screen "P_GraphicView_1" 1280x800
   GraphicView "Default" at 10,10 size 100x60
   TextField "Label_Default" at 10,72 size 108x16; Text 'Default'
   GraphicView "BackColor" at 120,10 size 100x60
   TextField "Label_BackColor" at 120,72 size 108x16; Text 'BackColor'
   GraphicView "BackFillStyle" at 230,10 size 100x60
   TextField "Label_BackFillStyle" at 230,72 size 108x16; Text 'BackFillStyle'
   GraphicView "BorderColor" at 340,10 size 100x60
   TextField "Label_BorderColor" at 340,72 size 108x16; Text 'BorderColor'
   GraphicView "BorderWidth" at 450,10 size 100x60
   TextField "Label_BorderWidth" at 450,72 size 108x16; Text 'BorderWidth'
   GraphicView "EdgeStyle" at 560,10 size 100x60
   TextField "Label_EdgeStyle" at 560,72 size 108x16; Text 'EdgeStyle'
   GraphicView "EdgeStyle_2" at 670,10 size 100x60
   TextField "Label_EdgeStyle_2" at 670,72 size 108x16; Text 'EdgeStyle_2'
   GraphicView "EdgeStyle_3" at 780,10 size 100x60
   TextField "Label_EdgeStyle_3" at 780,72 size 108x16; Text 'EdgeStyle_3'
   GraphicView "EdgeStyle_4" at 890,10 size 100x60
   TextField "Label_EdgeStyle_4" at 890,72 size 108x16; Text 'EdgeStyle_4'
   GraphicView "FitToLargest" at 1000,10 size 100x60
   TextField "Label_FitToLargest" at 1000,72 size 108x16; Text 'FitToLargest'
   GraphicView "Flashing" at 1110,10 size 100x60
   TextField "Label_Flashing" at 1110,72 size 108x16; Text 'Flashing'
   GraphicView "TransparentColor" at 10,96 size 100x60
   TextField "Label_TransparentColor" at 10,158 size 108x16; Text 'TransparentColor'
   GraphicView "UseTransparentColor" at 120,96 size 100x60
   TextField "Label_UseTransparentColor" at 120,158 size 108x16; Text 'UseTransparentColor'
   Button "Next" at 1238,776 size 40x22; TextOff 'Text'
      on Click: ActivateScreen("P_IOField_1", 0)

screen "P_IOField_1" 1280x800
   IOField "Default" at 10,10 size 100x30
   TextField "Label_Default" at 10,42 size 108x16; Text 'Default'
   IOField "AboveUpperLimitColor" at 120,10 size 100x30
   TextField "Label_AboveUpperLimitColor" at 120,42 size 108x16; Text 'AboveUpperLimitColor'
   IOField "BackColor" at 230,10 size 100x30
   TextField "Label_BackColor" at 230,42 size 108x16; Text 'BackColor'
   IOField "BackFillStyle" at 340,10 size 100x30
   TextField "Label_BackFillStyle" at 340,42 size 108x16; Text 'BackFillStyle'
   IOField "BelowLowerLimitColor" at 450,10 size 100x30
   TextField "Label_BelowLowerLimitColor" at 450,42 size 108x16; Text 'BelowLowerLimitColor'
   IOField "BorderBackColor" at 560,10 size 100x30
   TextField "Label_BorderBackColor" at 560,42 size 108x16; Text 'BorderBackColor'
   IOField "BorderColor" at 670,10 size 100x30
   TextField "Label_BorderColor" at 670,42 size 108x16; Text 'BorderColor'
   IOField "BorderWidth" at 780,10 size 100x30
   TextField "Label_BorderWidth" at 780,42 size 108x16; Text 'BorderWidth'
   IOField "BottomMargin" at 890,10 size 100x30
   TextField "Label_BottomMargin" at 890,42 size 108x16; Text 'BottomMargin'
   IOField "CornerRadius" at 1000,10 size 100x30
   TextField "Label_CornerRadius" at 1000,42 size 108x16; Text 'CornerRadius'
   IOField "DataFormat_3" at 1110,10 size 100x30
   TextField "Label_DataFormat_3" at 1110,42 size 108x16; Text 'DataFormat_3'
   IOField "EdgeStyle" at 10,66 size 100x30
   TextField "Label_EdgeStyle" at 10,98 size 108x16; Text 'EdgeStyle'
   IOField "EdgeStyle_2" at 120,66 size 100x30
   TextField "Label_EdgeStyle_2" at 120,98 size 108x16; Text 'EdgeStyle_2'
   IOField "EdgeStyle_3" at 230,66 size 100x30
   TextField "Label_EdgeStyle_3" at 230,98 size 108x16; Text 'EdgeStyle_3'
   IOField "EdgeStyle_4" at 340,66 size 100x30
   TextField "Label_EdgeStyle_4" at 340,98 size 108x16; Text 'EdgeStyle_4'
   IOField "FieldLength" at 450,66 size 100x30
   TextField "Label_FieldLength" at 450,98 size 108x16; Text 'FieldLength'
   IOField "FitToLargest" at 560,66 size 100x30
   TextField "Label_FitToLargest" at 560,98 size 108x16; Text 'FitToLargest'
   IOField "Flashing" at 670,66 size 100x30
   TextField "Label_Flashing" at 670,98 size 108x16; Text 'Flashing'
   IOField "ForeColor" at 780,66 size 100x30
   TextField "Label_ForeColor" at 780,98 size 108x16; Text 'ForeColor'
   IOField "FormatPattern" at 890,66 size 100x30; FormatPattern 99.9
   TextField "Label_FormatPattern" at 890,98 size 108x16; Text 'FormatPattern'
   IOField "HorizontalAlignment" at 1000,66 size 100x30
   TextField "Label_HorizontalAlignment" at 1000,98 size 108x16; Text 'HorizontalAlignment'
   IOField "HorizontalAlignment_2" at 1110,66 size 100x30
   TextField "Label_HorizontalAlignment_2" at 1110,98 size 108x16; Text 'HorizontalAlignment_2'
   IOField "LeftMargin" at 10,122 size 100x30
   TextField "Label_LeftMargin" at 10,154 size 108x16; Text 'LeftMargin'
   IOField "Mode" at 120,122 size 100x30
   TextField "Label_Mode" at 120,154 size 108x16; Text 'Mode'
   IOField "Mode_2" at 230,122 size 100x30
   TextField "Label_Mode_2" at 230,154 size 108x16; Text 'Mode_2'
   IOField "RightMargin" at 340,122 size 100x30
   TextField "Label_RightMargin" at 340,154 size 108x16; Text 'RightMargin'
   IOField "ShiftDecimalPoint" at 450,122 size 100x30
   TextField "Label_ShiftDecimalPoint" at 450,154 size 108x16; Text 'ShiftDecimalPoint'
   IOField "ShowLeadingZeros" at 560,122 size 100x30
   TextField "Label_ShowLeadingZeros" at 560,154 size 108x16; Text 'ShowLeadingZeros'
   IOField "TopMargin" at 670,122 size 100x30
   TextField "Label_TopMargin" at 670,154 size 108x16; Text 'TopMargin'
   IOField "Unit" at 780,122 size 100x30; Unit mm
   TextField "Label_Unit" at 780,154 size 108x16; Text 'Unit'
   IOField "UseDesignColorSchema" at 890,122 size 100x30
   TextField "Label_UseDesignColorSchema" at 890,154 size 108x16; Text 'UseDesignColorSchema'
   IOField "VerticalAlignment" at 1000,122 size 100x30
   TextField "Label_VerticalAlignment" at 1000,154 size 108x16; Text 'VerticalAlignment'
   IOField "VerticalAlignment_2" at 1110,122 size 100x30
   TextField "Label_VerticalAlignment_2" at 1110,154 size 108x16; Text 'VerticalAlignment_2'
   Button "Next" at 1238,776 size 40x22; TextOff 'Text'
      on Click: ActivateScreen("P_Button_1", 0)

screen "P_Button_1" 1280x800
   Button "Default" at 10,10 size 100x40; TextOff 'Text'
   TextField "Label_Default" at 10,52 size 108x16; Text 'Default'
   Button "BackColor" at 120,10 size 100x40; TextOff 'Text'
   TextField "Label_BackColor" at 120,52 size 108x16; Text 'BackColor'
   Button "BackFillStyle" at 230,10 size 100x40; TextOff 'Text'
   TextField "Label_BackFillStyle" at 230,52 size 108x16; Text 'BackFillStyle'
   Button "BorderBackColor" at 340,10 size 100x40; TextOff 'Text'
   TextField "Label_BorderBackColor" at 340,52 size 108x16; Text 'BorderBackColor'
   Button "BorderColor" at 450,10 size 100x40; TextOff 'Text'
   TextField "Label_BorderColor" at 450,52 size 108x16; Text 'BorderColor'
   Button "BorderWidth" at 560,10 size 100x40; TextOff 'Text'
   TextField "Label_BorderWidth" at 560,52 size 108x16; Text 'BorderWidth'
   Button "CornerRadius" at 670,10 size 100x40; TextOff 'Text'
   TextField "Label_CornerRadius" at 670,52 size 108x16; Text 'CornerRadius'
   Button "EdgeStyle" at 780,10 size 100x40; TextOff 'Text'
   TextField "Label_EdgeStyle" at 780,52 size 108x16; Text 'EdgeStyle'
   Button "EdgeStyle_2" at 890,10 size 100x40; TextOff 'Text'
   TextField "Label_EdgeStyle_2" at 890,52 size 108x16; Text 'EdgeStyle_2'
   Button "EdgeStyle_3" at 1000,10 size 100x40; TextOff 'Text'
   TextField "Label_EdgeStyle_3" at 1000,52 size 108x16; Text 'EdgeStyle_3'
   Button "EdgeStyle_4" at 1110,10 size 100x40; TextOff 'Text'
   TextField "Label_EdgeStyle_4" at 1110,52 size 108x16; Text 'EdgeStyle_4'
   Button "FirstGradientColor" at 10,76 size 100x40; TextOff 'Text'
   TextField "Label_FirstGradientColor" at 10,118 size 108x16; Text 'FirstGradientColor'
   Button "FirstGradientOffset" at 120,76 size 100x40; TextOff 'Text'
   TextField "Label_FirstGradientOffset" at 120,118 size 108x16; Text 'FirstGradientOffset'
   Button "FitToLargest" at 230,76 size 100x40; TextOff 'Text'
   TextField "Label_FitToLargest" at 230,118 size 108x16; Text 'FitToLargest'
   Button "Flashing" at 340,76 size 100x40; TextOff 'Text'
   TextField "Label_Flashing" at 340,118 size 108x16; Text 'Flashing'
   Button "FocusColor" at 450,76 size 100x40; TextOff 'Text'
   TextField "Label_FocusColor" at 450,118 size 108x16; Text 'FocusColor'
   Button "FocusWidth" at 560,76 size 100x40; TextOff 'Text'
   TextField "Label_FocusWidth" at 560,118 size 108x16; Text 'FocusWidth'
   Button "ForeColor" at 670,76 size 100x40; TextOff 'Text'
   TextField "Label_ForeColor" at 670,118 size 108x16; Text 'ForeColor'
   Button "HorizontalAlignment" at 780,76 size 100x40; TextOff 'Text'
   TextField "Label_HorizontalAlignment" at 780,118 size 108x16; Text 'HorizontalAlignment'
   Button "HorizontalAlignment_2" at 890,76 size 100x40; TextOff 'Text'
   TextField "Label_HorizontalAlignment_2" at 890,118 size 108x16; Text 'HorizontalAlignment_2'
   Button "HorizontalPictureAlignment" at 1000,76 size 100x40; TextOff 'Text'
   TextField "Label_HorizontalPictureAlignment" at 1000,118 size 108x16; Text 'HorizontalPictureAlignment'
   Button "HorizontalPictureAlignment_2" at 1110,76 size 100x40; TextOff 'Text'
   TextField "Label_HorizontalPictureAlignment_2" at 1110,118 size 108x16; Text 'HorizontalPictureAlignment_2'
   Button "MiddleGradientColor" at 10,142 size 100x40; TextOff 'Text'
   TextField "Label_MiddleGradientColor" at 10,184 size 108x16; Text 'MiddleGradientColor'
   Button "Mode_5" at 120,142 size 100x40; TextOff 'Text'
   TextField "Label_Mode_5" at 120,184 size 108x16; Text 'Mode_5'
   Button "Mode_7" at 230,142 size 100x40; TextOff 'Text'
   TextField "Label_Mode_7" at 230,184 size 108x16; Text 'Mode_7'
   Button "PictureAreaBottomMargin" at 340,142 size 100x40; TextOff 'Text'
   TextField "Label_PictureAreaBottomMargin" at 340,184 size 108x16; Text 'PictureAreaBottomMargin'
   Button "PictureAreaLeftMargin" at 450,142 size 100x40; TextOff 'Text'
   TextField "Label_PictureAreaLeftMargin" at 450,184 size 108x16; Text 'PictureAreaLeftMargin'
   Button "PictureAreaRightMargin" at 560,142 size 100x40; TextOff 'Text'
   TextField "Label_PictureAreaRightMargin" at 560,184 size 108x16; Text 'PictureAreaRightMargin'
   Button "PictureAreaTopMargin" at 670,142 size 100x40; TextOff 'Text'
   TextField "Label_PictureAreaTopMargin" at 670,184 size 108x16; Text 'PictureAreaTopMargin'
   Button "SecondGradientColor" at 780,142 size 100x40; TextOff 'Text'
   TextField "Label_SecondGradientColor" at 780,184 size 108x16; Text 'SecondGradientColor'
   Button "SecondGradientOffset" at 890,142 size 100x40; TextOff 'Text'
   TextField "Label_SecondGradientOffset" at 890,184 size 108x16; Text 'SecondGradientOffset'
   Button "TextAreaBottomMargin" at 1000,142 size 100x40; TextOff 'Text'
   TextField "Label_TextAreaBottomMargin" at 1000,184 size 108x16; Text 'TextAreaBottomMargin'
   Button "TextAreaLeftMargin" at 1110,142 size 100x40; TextOff 'Text'
   TextField "Label_TextAreaLeftMargin" at 1110,184 size 108x16; Text 'TextAreaLeftMargin'
   Button "TextAreaRightMargin" at 10,208 size 100x40; TextOff 'Text'
   TextField "Label_TextAreaRightMargin" at 10,250 size 108x16; Text 'TextAreaRightMargin'
   Button "TextAreaTopMargin" at 120,208 size 100x40; TextOff 'Text'
   TextField "Label_TextAreaTopMargin" at 120,250 size 108x16; Text 'TextAreaTopMargin'
   Button "UseDesignColorSchema" at 230,208 size 100x40; TextOff 'Text'
   TextField "Label_UseDesignColorSchema" at 230,250 size 108x16; Text 'UseDesignColorSchema'
   Button "UseFirstGradient" at 340,208 size 100x40; TextOff 'Text'
   TextField "Label_UseFirstGradient" at 340,250 size 108x16; Text 'UseFirstGradient'
   Button "UseSecondGradient" at 450,208 size 100x40; TextOff 'Text'
   TextField "Label_UseSecondGradient" at 450,250 size 108x16; Text 'UseSecondGradient'
   Button "VerticalAlignment" at 560,208 size 100x40; TextOff 'Text'
   TextField "Label_VerticalAlignment" at 560,250 size 108x16; Text 'VerticalAlignment'
   Button "VerticalAlignment_2" at 670,208 size 100x40; TextOff 'Text'
   TextField "Label_VerticalAlignment_2" at 670,250 size 108x16; Text 'VerticalAlignment_2'
   Button "VerticalPictureAlignment" at 780,208 size 100x40; TextOff 'Text'
   TextField "Label_VerticalPictureAlignment" at 780,250 size 108x16; Text 'VerticalPictureAlignment'
   Button "VerticalPictureAlignment_2" at 890,208 size 100x40; TextOff 'Text'
   TextField "Label_VerticalPictureAlignment_2" at 890,250 size 108x16; Text 'VerticalPictureAlignment_2'
   Button "Next" at 1238,776 size 40x22; TextOff 'Text'
      on Click: ActivateScreen("P_SymbolicIOField_1", 0)

screen "P_SymbolicIOField_1" 1280x800
   SymbolicIOField "Default" at 10,10 size 120x30; TextOff '0'; TextOn '1'
   TextField "Label_Default" at 10,42 size 128x16; Text 'Default'
   SymbolicIOField "AboveUpperLimitColor" at 140,10 size 120x30; TextOff '0'; TextOn '1'
   TextField "Label_AboveUpperLimitColor" at 140,42 size 128x16; Text 'AboveUpperLimitColor'
   SymbolicIOField "BackColor" at 270,10 size 120x30; TextOff '0'; TextOn '1'
   TextField "Label_BackColor" at 270,42 size 128x16; Text 'BackColor'
   SymbolicIOField "BackFillStyle" at 400,10 size 120x30; TextOff '0'; TextOn '1'
   TextField "Label_BackFillStyle" at 400,42 size 128x16; Text 'BackFillStyle'
   SymbolicIOField "BelowLowerLimitColor" at 530,10 size 120x30; TextOff '0'; TextOn '1'
   TextField "Label_BelowLowerLimitColor" at 530,42 size 128x16; Text 'BelowLowerLimitColor'
   SymbolicIOField "BorderBackColor" at 660,10 size 120x30; TextOff '0'; TextOn '1'
   TextField "Label_BorderBackColor" at 660,42 size 128x16; Text 'BorderBackColor'
   SymbolicIOField "BorderColor" at 790,10 size 120x30; TextOff '0'; TextOn '1'
   TextField "Label_BorderColor" at 790,42 size 128x16; Text 'BorderColor'
   SymbolicIOField "BorderWidth" at 920,10 size 120x30; TextOff '0'; TextOn '1'
   TextField "Label_BorderWidth" at 920,42 size 128x16; Text 'BorderWidth'
   SymbolicIOField "BottomMargin" at 1050,10 size 120x30; TextOff '0'; TextOn '1'
   TextField "Label_BottomMargin" at 1050,42 size 128x16; Text 'BottomMargin'
   SymbolicIOField "CornerRadius" at 10,66 size 120x30; TextOff '0'; TextOn '1'
   TextField "Label_CornerRadius" at 10,98 size 128x16; Text 'CornerRadius'
   SymbolicIOField "CountVisibleItems" at 140,66 size 120x30; TextOff '0'; TextOn '1'
   TextField "Label_CountVisibleItems" at 140,98 size 128x16; Text 'CountVisibleItems'
   SymbolicIOField "EdgeStyle" at 270,66 size 120x30; TextOff '0'; TextOn '1'
   TextField "Label_EdgeStyle" at 270,98 size 128x16; Text 'EdgeStyle'
   SymbolicIOField "EdgeStyle_2" at 400,66 size 120x30; TextOff '0'; TextOn '1'
   TextField "Label_EdgeStyle_2" at 400,98 size 128x16; Text 'EdgeStyle_2'
   SymbolicIOField "EdgeStyle_3" at 530,66 size 120x30; TextOff '0'; TextOn '1'
   TextField "Label_EdgeStyle_3" at 530,98 size 128x16; Text 'EdgeStyle_3'
   SymbolicIOField "EdgeStyle_4" at 660,66 size 120x30; TextOff '0'; TextOn '1'
   TextField "Label_EdgeStyle_4" at 660,98 size 128x16; Text 'EdgeStyle_4'
   SymbolicIOField "EvenRowBackColor" at 790,66 size 120x30; TextOff '0'; TextOn '1'
   TextField "Label_EvenRowBackColor" at 790,98 size 128x16; Text 'EvenRowBackColor'
   SymbolicIOField "FitToLargest" at 920,66 size 120x30; TextOff '0'; TextOn '1'
   TextField "Label_FitToLargest" at 920,98 size 128x16; Text 'FitToLargest'
   SymbolicIOField "Flashing" at 1050,66 size 120x30; TextOff '0'; TextOn '1'
   TextField "Label_Flashing" at 1050,98 size 128x16; Text 'Flashing'
   SymbolicIOField "FlashingOnLimitViolation" at 10,122 size 120x30; TextOff '0'; TextOn '1'
   TextField "Label_FlashingOnLimitViolation" at 10,154 size 128x16; Text 'FlashingOnLimitViolation'
   SymbolicIOField "ForeColor" at 140,122 size 120x30; TextOff '0'; TextOn '1'
   TextField "Label_ForeColor" at 140,154 size 128x16; Text 'ForeColor'
   SymbolicIOField "HorizontalAlignment" at 270,122 size 120x30; TextOff '0'; TextOn '1'
   TextField "Label_HorizontalAlignment" at 270,154 size 128x16; Text 'HorizontalAlignment'
   SymbolicIOField "HorizontalAlignment_2" at 400,122 size 120x30; TextOff '0'; TextOn '1'
   TextField "Label_HorizontalAlignment_2" at 400,154 size 128x16; Text 'HorizontalAlignment_2'
   SymbolicIOField "LeftMargin" at 530,122 size 120x30; TextOff '0'; TextOn '1'
   TextField "Label_LeftMargin" at 530,154 size 128x16; Text 'LeftMargin'
   SymbolicIOField "Mode" at 660,122 size 120x30; TextOff '0'; TextOn '1'
   TextField "Label_Mode" at 660,154 size 128x16; Text 'Mode'
   SymbolicIOField "Mode_2" at 790,122 size 120x30; TextOff '0'; TextOn '1'
   TextField "Label_Mode_2" at 790,154 size 128x16; Text 'Mode_2'
   SymbolicIOField "RightMargin" at 920,122 size 120x30; TextOff '0'; TextOn '1'
   TextField "Label_RightMargin" at 920,154 size 128x16; Text 'RightMargin'
   SymbolicIOField "SelectBackColor" at 1050,122 size 120x30; TextOff '0'; TextOn '1'
   TextField "Label_SelectBackColor" at 1050,154 size 128x16; Text 'SelectBackColor'
   SymbolicIOField "SelectForeColor" at 10,178 size 120x30; TextOff '0'; TextOn '1'
   TextField "Label_SelectForeColor" at 10,210 size 128x16; Text 'SelectForeColor'
   SymbolicIOField "ShowDropDownButton" at 140,178 size 120x30; TextOff '0'; TextOn '1'
   TextField "Label_ShowDropDownButton" at 140,210 size 128x16; Text 'ShowDropDownButton'
   SymbolicIOField "ShowDropDownList" at 270,178 size 120x30; TextOff '0'; TextOn '1'
   TextField "Label_ShowDropDownList" at 270,210 size 128x16; Text 'ShowDropDownList'
   SymbolicIOField "TopMargin" at 400,178 size 120x30; TextOff '0'; TextOn '1'
   TextField "Label_TopMargin" at 400,210 size 128x16; Text 'TopMargin'
   SymbolicIOField "UseDesignColorSchema" at 530,178 size 120x30; TextOff '0'; TextOn '1'
   TextField "Label_UseDesignColorSchema" at 530,210 size 128x16; Text 'UseDesignColorSchema'
   SymbolicIOField "VerticalAlignment" at 660,178 size 120x30; TextOff '0'; TextOn '1'
   TextField "Label_VerticalAlignment" at 660,210 size 128x16; Text 'VerticalAlignment'
   SymbolicIOField "VerticalAlignment_2" at 790,178 size 120x30; TextOff '0'; TextOn '1'
   TextField "Label_VerticalAlignment_2" at 790,210 size 128x16; Text 'VerticalAlignment_2'
   Button "Next" at 1238,776 size 40x22; TextOff 'Text'
      on Click: ActivateScreen("P_GraphicIOField_1", 0)

screen "P_GraphicIOField_1" 1280x800
   GraphicIOField "Default" at 10,10 size 60x60
   TextField "Label_Default" at 10,72 size 68x16; Text 'Default'
   GraphicIOField "AboveUpperLimitColor" at 80,10 size 60x60
   TextField "Label_AboveUpperLimitColor" at 80,72 size 68x16; Text 'AboveUpperLimitColor'
   GraphicIOField "BackColor" at 150,10 size 60x60
   TextField "Label_BackColor" at 150,72 size 68x16; Text 'BackColor'
   GraphicIOField "BackFillStyle" at 220,10 size 60x60
   TextField "Label_BackFillStyle" at 220,72 size 68x16; Text 'BackFillStyle'
   GraphicIOField "BelowLowerLimitColor" at 290,10 size 60x60
   TextField "Label_BelowLowerLimitColor" at 290,72 size 68x16; Text 'BelowLowerLimitColor'
   GraphicIOField "BorderColor" at 360,10 size 60x60
   TextField "Label_BorderColor" at 360,72 size 68x16; Text 'BorderColor'
   GraphicIOField "BorderWidth" at 430,10 size 60x60
   TextField "Label_BorderWidth" at 430,72 size 68x16; Text 'BorderWidth'
   GraphicIOField "EdgeStyle" at 500,10 size 60x60
   TextField "Label_EdgeStyle" at 500,72 size 68x16; Text 'EdgeStyle'
   GraphicIOField "EdgeStyle_2" at 570,10 size 60x60
   TextField "Label_EdgeStyle_2" at 570,72 size 68x16; Text 'EdgeStyle_2'
   GraphicIOField "EdgeStyle_3" at 640,10 size 60x60
   TextField "Label_EdgeStyle_3" at 640,72 size 68x16; Text 'EdgeStyle_3'
   GraphicIOField "EdgeStyle_4" at 710,10 size 60x60
   TextField "Label_EdgeStyle_4" at 710,72 size 68x16; Text 'EdgeStyle_4'
   GraphicIOField "FitToLargest" at 780,10 size 60x60
   TextField "Label_FitToLargest" at 780,72 size 68x16; Text 'FitToLargest'
   GraphicIOField "Flashing" at 850,10 size 60x60
   TextField "Label_Flashing" at 850,72 size 68x16; Text 'Flashing'
   GraphicIOField "FlashingOnLimitViolation" at 920,10 size 60x60
   TextField "Label_FlashingOnLimitViolation" at 920,72 size 68x16; Text 'FlashingOnLimitViolation'
   GraphicIOField "FocusColor" at 990,10 size 60x60
   TextField "Label_FocusColor" at 990,72 size 68x16; Text 'FocusColor'
   GraphicIOField "FocusWidth" at 1060,10 size 60x60
   TextField "Label_FocusWidth" at 1060,72 size 68x16; Text 'FocusWidth'
   GraphicIOField "Mode" at 1130,10 size 60x60
   TextField "Label_Mode" at 1130,72 size 68x16; Text 'Mode'
   GraphicIOField "Mode_2" at 1200,10 size 60x60
   TextField "Label_Mode_2" at 1200,72 size 68x16; Text 'Mode_2'
   GraphicIOField "ScrollBarOrientation" at 10,96 size 60x60
   TextField "Label_ScrollBarOrientation" at 10,158 size 68x16; Text 'ScrollBarOrientation'
   GraphicIOField "TransparentColor" at 80,96 size 60x60
   TextField "Label_TransparentColor" at 80,158 size 68x16; Text 'TransparentColor'
   GraphicIOField "UseTransparentColor" at 150,96 size 60x60
   TextField "Label_UseTransparentColor" at 150,158 size 68x16; Text 'UseTransparentColor'
   Button "Next" at 1238,776 size 40x22; TextOff 'Text'
      on Click: ActivateScreen("P_DateTimeField_1", 0)

screen "P_DateTimeField_1" 1280x800
   DateTimeField "Default" at 10,10 size 160x30
   TextField "Label_Default" at 10,42 size 168x16; Text 'Default'
   DateTimeField "BackColor" at 180,10 size 160x30
   TextField "Label_BackColor" at 180,42 size 168x16; Text 'BackColor'
   DateTimeField "BackFillStyle" at 350,10 size 160x30
   TextField "Label_BackFillStyle" at 350,42 size 168x16; Text 'BackFillStyle'
   DateTimeField "BorderBackColor" at 520,10 size 160x30
   TextField "Label_BorderBackColor" at 520,42 size 168x16; Text 'BorderBackColor'
   DateTimeField "BorderColor" at 690,10 size 160x30
   TextField "Label_BorderColor" at 690,42 size 168x16; Text 'BorderColor'
   DateTimeField "BorderWidth" at 860,10 size 160x30
   TextField "Label_BorderWidth" at 860,42 size 168x16; Text 'BorderWidth'
   DateTimeField "BottomMargin" at 1030,10 size 160x30
   TextField "Label_BottomMargin" at 1030,42 size 168x16; Text 'BottomMargin'
   DateTimeField "CornerRadius" at 10,66 size 160x30
   TextField "Label_CornerRadius" at 10,98 size 168x16; Text 'CornerRadius'
   DateTimeField "DisplaySystemTime" at 180,66 size 160x30
   TextField "Label_DisplaySystemTime" at 180,98 size 168x16; Text 'DisplaySystemTime'
   DateTimeField "EdgeStyle" at 350,66 size 160x30
   TextField "Label_EdgeStyle" at 350,98 size 168x16; Text 'EdgeStyle'
   DateTimeField "EdgeStyle_2" at 520,66 size 160x30
   TextField "Label_EdgeStyle_2" at 520,98 size 168x16; Text 'EdgeStyle_2'
   DateTimeField "EdgeStyle_3" at 690,66 size 160x30
   TextField "Label_EdgeStyle_3" at 690,98 size 168x16; Text 'EdgeStyle_3'
   DateTimeField "EdgeStyle_4" at 860,66 size 160x30
   TextField "Label_EdgeStyle_4" at 860,98 size 168x16; Text 'EdgeStyle_4'
   DateTimeField "FitToLargest" at 1030,66 size 160x30
   TextField "Label_FitToLargest" at 1030,98 size 168x16; Text 'FitToLargest'
   DateTimeField "Flashing" at 10,122 size 160x30
   TextField "Label_Flashing" at 10,154 size 168x16; Text 'Flashing'
   DateTimeField "ForeColor" at 180,122 size 160x30
   TextField "Label_ForeColor" at 180,154 size 168x16; Text 'ForeColor'
   DateTimeField "HorizontalAlignment" at 350,122 size 160x30
   TextField "Label_HorizontalAlignment" at 350,154 size 168x16; Text 'HorizontalAlignment'
   DateTimeField "HorizontalAlignment_2" at 520,122 size 160x30
   TextField "Label_HorizontalAlignment_2" at 520,154 size 168x16; Text 'HorizontalAlignment_2'
   DateTimeField "LeftMargin" at 690,122 size 160x30
   TextField "Label_LeftMargin" at 690,154 size 168x16; Text 'LeftMargin'
   DateTimeField "LongDateTimeFormat" at 860,122 size 160x30
   TextField "Label_LongDateTimeFormat" at 860,154 size 168x16; Text 'LongDateTimeFormat'
   DateTimeField "Mode_3" at 1030,122 size 160x30
   TextField "Label_Mode_3" at 1030,154 size 168x16; Text 'Mode_3'
   DateTimeField "RightMargin" at 10,178 size 160x30
   TextField "Label_RightMargin" at 10,210 size 168x16; Text 'RightMargin'
   DateTimeField "ShowDate" at 180,178 size 160x30
   TextField "Label_ShowDate" at 180,210 size 168x16; Text 'ShowDate'
   DateTimeField "ShowTime" at 350,178 size 160x30
   TextField "Label_ShowTime" at 350,210 size 168x16; Text 'ShowTime'
   DateTimeField "TopMargin" at 520,178 size 160x30
   TextField "Label_TopMargin" at 520,210 size 168x16; Text 'TopMargin'
   DateTimeField "UseDesignColorSchema" at 690,178 size 160x30
   TextField "Label_UseDesignColorSchema" at 690,210 size 168x16; Text 'UseDesignColorSchema'
   DateTimeField "VerticalAlignment" at 860,178 size 160x30
   TextField "Label_VerticalAlignment" at 860,210 size 168x16; Text 'VerticalAlignment'
   DateTimeField "VerticalAlignment_2" at 1030,178 size 160x30
   TextField "Label_VerticalAlignment_2" at 1030,210 size 168x16; Text 'VerticalAlignment_2'
   Button "Next" at 1238,776 size 40x22; TextOff 'Text'
      on Click: ActivateScreen("P_Bar_1", 0)

screen "P_Bar_1" 1280x800
   Bar "Default" at 10,10 size 40x120
   TextField "Label_Default" at 10,132 size 48x16; Text 'Default'
   Bar "BackColor" at 60,10 size 40x120
   TextField "Label_BackColor" at 60,132 size 48x16; Text 'BackColor'
   Bar "BarBackColor" at 110,10 size 40x120
   TextField "Label_BarBackColor" at 110,132 size 48x16; Text 'BarBackColor'
   Bar "BarEdgeStyle" at 160,10 size 40x120
   TextField "Label_BarEdgeStyle" at 160,132 size 48x16; Text 'BarEdgeStyle'
   Bar "BarEdgeStyle_2" at 210,10 size 40x120
   TextField "Label_BarEdgeStyle_2" at 210,132 size 48x16; Text 'BarEdgeStyle_2'
   Bar "BarOrientation" at 260,10 size 40x120
   TextField "Label_BarOrientation" at 260,132 size 48x16; Text 'BarOrientation'
   Bar "BarOrientation_2" at 310,10 size 40x120
   TextField "Label_BarOrientation_2" at 310,132 size 48x16; Text 'BarOrientation_2'
   Bar "BarOrientation_3" at 360,10 size 40x120
   TextField "Label_BarOrientation_3" at 360,132 size 48x16; Text 'BarOrientation_3'
   Bar "BorderBackColor" at 410,10 size 40x120
   TextField "Label_BorderBackColor" at 410,132 size 48x16; Text 'BorderBackColor'
   Bar "BorderColor" at 460,10 size 40x120
   TextField "Label_BorderColor" at 460,132 size 48x16; Text 'BorderColor'
   Bar "BorderWidth" at 510,10 size 40x120
   TextField "Label_BorderWidth" at 510,132 size 48x16; Text 'BorderWidth'
   Bar "CornerRadius" at 560,10 size 40x120
   TextField "Label_CornerRadius" at 560,132 size 48x16; Text 'CornerRadius'
   Bar "CountSubDivisions" at 610,10 size 40x120
   TextField "Label_CountSubDivisions" at 610,132 size 48x16; Text 'CountSubDivisions'
   Bar "EdgeStyle" at 660,10 size 40x120
   TextField "Label_EdgeStyle" at 660,132 size 48x16; Text 'EdgeStyle'
   Bar "EdgeStyle_2" at 710,10 size 40x120
   TextField "Label_EdgeStyle_2" at 710,132 size 48x16; Text 'EdgeStyle_2'
   Bar "EdgeStyle_3" at 760,10 size 40x120
   TextField "Label_EdgeStyle_3" at 760,132 size 48x16; Text 'EdgeStyle_3'
   Bar "EdgeStyle_4" at 810,10 size 40x120
   TextField "Label_EdgeStyle_4" at 810,132 size 48x16; Text 'EdgeStyle_4'
   Bar "Flashing" at 860,10 size 40x120
   TextField "Label_Flashing" at 860,132 size 48x16; Text 'Flashing'
   Bar "FlashingOnLimitViolation" at 910,10 size 40x120
   TextField "Label_FlashingOnLimitViolation" at 910,132 size 48x16; Text 'FlashingOnLimitViolation'
   Bar "ForeColor" at 960,10 size 40x120
   TextField "Label_ForeColor" at 960,132 size 48x16; Text 'ForeColor'
   Bar "IntegerDigits" at 1010,10 size 40x120
   TextField "Label_IntegerDigits" at 1010,132 size 48x16; Text 'IntegerDigits'
   Bar "LargeTickLabelingStep" at 1060,10 size 40x120
   TextField "Label_LargeTickLabelingStep" at 1060,132 size 48x16; Text 'LargeTickLabelingStep'
   Bar "MaximumValue" at 1110,10 size 40x120; MaximumValue 200
   TextField "Label_MaximumValue" at 1110,132 size 48x16; Text 'MaximumValue'
   Bar "MinimumValue" at 1160,10 size 40x120; MinimumValue -100
   TextField "Label_MinimumValue" at 1160,132 size 48x16; Text 'MinimumValue'
   Bar "Precision" at 1210,10 size 40x120
   TextField "Label_Precision" at 1210,132 size 48x16; Text 'Precision'
   Bar "RangeLower1Color" at 10,156 size 40x120
   TextField "Label_RangeLower1Color" at 10,278 size 48x16; Text 'RangeLower1Color'
   Bar "RangeLower1Enabled" at 60,156 size 40x120
   TextField "Label_RangeLower1Enabled" at 60,278 size 48x16; Text 'RangeLower1Enabled'
   Bar "RangeLower2Color" at 110,156 size 40x120
   TextField "Label_RangeLower2Color" at 110,278 size 48x16; Text 'RangeLower2Color'
   Bar "RangeLower2Enabled" at 160,156 size 40x120
   TextField "Label_RangeLower2Enabled" at 160,278 size 48x16; Text 'RangeLower2Enabled'
   Bar "RangeNormalColor" at 210,156 size 40x120
   TextField "Label_RangeNormalColor" at 210,278 size 48x16; Text 'RangeNormalColor'
   Bar "RangeNormalEnabled" at 260,156 size 40x120
   TextField "Label_RangeNormalEnabled" at 260,278 size 48x16; Text 'RangeNormalEnabled'
   Bar "RangeUpper1Color" at 310,156 size 40x120
   TextField "Label_RangeUpper1Color" at 310,278 size 48x16; Text 'RangeUpper1Color'
   Bar "RangeUpper1Enabled" at 360,156 size 40x120
   TextField "Label_RangeUpper1Enabled" at 360,278 size 48x16; Text 'RangeUpper1Enabled'
   Bar "RangeUpper2Color" at 410,156 size 40x120
   TextField "Label_RangeUpper2Color" at 410,278 size 48x16; Text 'RangeUpper2Color'
   Bar "RangeUpper2Enabled" at 460,156 size 40x120
   TextField "Label_RangeUpper2Enabled" at 460,278 size 48x16; Text 'RangeUpper2Enabled'
   Bar "ScaleColor" at 510,156 size 40x120
   TextField "Label_ScaleColor" at 510,278 size 48x16; Text 'ScaleColor'
   Bar "ScaleGradation" at 560,156 size 40x120
   TextField "Label_ScaleGradation" at 560,278 size 48x16; Text 'ScaleGradation'
   Bar "ScaleLabelingDoubleLined" at 610,156 size 40x120
   TextField "Label_ScaleLabelingDoubleLined" at 610,278 size 48x16; Text 'ScaleLabelingDoubleLined'
   Bar "ScalePosition" at 660,156 size 40x120
   TextField "Label_ScalePosition" at 660,278 size 48x16; Text 'ScalePosition'
   Bar "SegmentColoring" at 710,156 size 40x120
   TextField "Label_SegmentColoring" at 710,278 size 48x16; Text 'SegmentColoring'
   Bar "ShowLimitLines" at 760,156 size 40x120
   TextField "Label_ShowLimitLines" at 760,278 size 48x16; Text 'ShowLimitLines'
   Bar "ShowLimitMarkers" at 810,156 size 40x120
   TextField "Label_ShowLimitMarkers" at 810,278 size 48x16; Text 'ShowLimitMarkers'
   Bar "ShowLimitRanges" at 860,156 size 40x120
   TextField "Label_ShowLimitRanges" at 860,278 size 48x16; Text 'ShowLimitRanges'
   Bar "ShowProcessValue" at 910,156 size 40x120
   TextField "Label_ShowProcessValue" at 910,278 size 48x16; Text 'ShowProcessValue'
   Bar "ShowScale" at 960,156 size 40x120
   TextField "Label_ShowScale" at 960,278 size 48x16; Text 'ShowScale'
   Bar "ShowTickLabels" at 1010,156 size 40x120
   TextField "Label_ShowTickLabels" at 1010,278 size 48x16; Text 'ShowTickLabels'
   Bar "Unit" at 1060,156 size 40x120; Unit mm
   TextField "Label_Unit" at 1060,278 size 48x16; Text 'Unit'
   Bar "UseAutoScaling" at 1110,156 size 40x120
   TextField "Label_UseAutoScaling" at 1110,278 size 48x16; Text 'UseAutoScaling'
   Bar "UseDesignColorSchema" at 1160,156 size 40x120
   TextField "Label_UseDesignColorSchema" at 1160,278 size 48x16; Text 'UseDesignColorSchema'
   Bar "UseExponentialFormat" at 1210,156 size 40x120
   TextField "Label_UseExponentialFormat" at 1210,278 size 48x16; Text 'UseExponentialFormat'
   Button "Next" at 1238,776 size 40x22; TextOff 'Text'
      on Click: ActivateScreen("P_Switch_1", 0)

screen "P_Switch_1" 1280x800
   Switch "Default" at 10,10 size 120x40; CaptionText 'Switch'; TextOff '0'; TextOn '1'
   TextField "Label_Default" at 10,52 size 128x16; Text 'Default'
   Switch "AboveUpperLimitColor" at 140,10 size 120x40; CaptionText 'Switch'; TextOff '0'; TextOn '1'
   TextField "Label_AboveUpperLimitColor" at 140,52 size 128x16; Text 'AboveUpperLimitColor'
   Switch "BackColor" at 270,10 size 120x40; CaptionText 'Switch'; TextOff '0'; TextOn '1'
   TextField "Label_BackColor" at 270,52 size 128x16; Text 'BackColor'
   Switch "BackFillStyle" at 400,10 size 120x40; CaptionText 'Switch'; TextOff '0'; TextOn '1'
   TextField "Label_BackFillStyle" at 400,52 size 128x16; Text 'BackFillStyle'
   Switch "BelowLowerLimitColor" at 530,10 size 120x40; CaptionText 'Switch'; TextOff '0'; TextOn '1'
   TextField "Label_BelowLowerLimitColor" at 530,52 size 128x16; Text 'BelowLowerLimitColor'
   Switch "BorderBackColor" at 660,10 size 120x40; CaptionText 'Switch'; TextOff '0'; TextOn '1'
   TextField "Label_BorderBackColor" at 660,52 size 128x16; Text 'BorderBackColor'
   Switch "BorderColor" at 790,10 size 120x40; CaptionText 'Switch'; TextOff '0'; TextOn '1'
   TextField "Label_BorderColor" at 790,52 size 128x16; Text 'BorderColor'
   Switch "BorderWidth" at 920,10 size 120x40; CaptionText 'Switch'; TextOff '0'; TextOn '1'
   TextField "Label_BorderWidth" at 920,52 size 128x16; Text 'BorderWidth'
   Switch "CaptionColor" at 1050,10 size 120x40; CaptionText 'Switch'; TextOff '0'; TextOn '1'
   TextField "Label_CaptionColor" at 1050,52 size 128x16; Text 'CaptionColor'
   Switch "CornerRadius" at 10,76 size 120x40; CaptionText 'Switch'; TextOff '0'; TextOn '1'
   TextField "Label_CornerRadius" at 10,118 size 128x16; Text 'CornerRadius'
   Switch "EdgeStyle" at 140,76 size 120x40; CaptionText 'Switch'; TextOff '0'; TextOn '1'
   TextField "Label_EdgeStyle" at 140,118 size 128x16; Text 'EdgeStyle'
   Switch "EdgeStyle_2" at 270,76 size 120x40; CaptionText 'Switch'; TextOff '0'; TextOn '1'
   TextField "Label_EdgeStyle_2" at 270,118 size 128x16; Text 'EdgeStyle_2'
   Switch "EdgeStyle_3" at 400,76 size 120x40; CaptionText 'Switch'; TextOff '0'; TextOn '1'
   TextField "Label_EdgeStyle_3" at 400,118 size 128x16; Text 'EdgeStyle_3'
   Switch "EdgeStyle_4" at 530,76 size 120x40; CaptionText 'Switch'; TextOff '0'; TextOn '1'
   TextField "Label_EdgeStyle_4" at 530,118 size 128x16; Text 'EdgeStyle_4'
   Switch "FirstGradientColor" at 660,76 size 120x40; CaptionText 'Switch'; TextOff '0'; TextOn '1'
   TextField "Label_FirstGradientColor" at 660,118 size 128x16; Text 'FirstGradientColor'
   Switch "FirstGradientOffset" at 790,76 size 120x40; CaptionText 'Switch'; TextOff '0'; TextOn '1'
   TextField "Label_FirstGradientOffset" at 790,118 size 128x16; Text 'FirstGradientOffset'
   Switch "FitToLargest" at 920,76 size 120x40; CaptionText 'Switch'; TextOff '0'; TextOn '1'
   TextField "Label_FitToLargest" at 920,118 size 128x16; Text 'FitToLargest'
   Switch "Flashing" at 1050,76 size 120x40; CaptionText 'Switch'; TextOff '0'; TextOn '1'
   TextField "Label_Flashing" at 1050,118 size 128x16; Text 'Flashing'
   Switch "FlashingOnLimitViolation" at 10,142 size 120x40; CaptionText 'Switch'; TextOff '0'; TextOn '1'
   TextField "Label_FlashingOnLimitViolation" at 10,184 size 128x16; Text 'FlashingOnLimitViolation'
   Switch "FocusColor" at 140,142 size 120x40; CaptionText 'Switch'; TextOff '0'; TextOn '1'
   TextField "Label_FocusColor" at 140,184 size 128x16; Text 'FocusColor'
   Switch "FocusWidth" at 270,142 size 120x40; CaptionText 'Switch'; TextOff '0'; TextOn '1'
   TextField "Label_FocusWidth" at 270,184 size 128x16; Text 'FocusWidth'
   Switch "ForeColor" at 400,142 size 120x40; CaptionText 'Switch'; TextOff '0'; TextOn '1'
   TextField "Label_ForeColor" at 400,184 size 128x16; Text 'ForeColor'
   Switch "HorizontalAlignment" at 530,142 size 120x40; CaptionText 'Switch'; TextOff '0'; TextOn '1'
   TextField "Label_HorizontalAlignment" at 530,184 size 128x16; Text 'HorizontalAlignment'
   Switch "HorizontalAlignment_2" at 660,142 size 120x40; CaptionText 'Switch'; TextOff '0'; TextOn '1'
   TextField "Label_HorizontalAlignment_2" at 660,184 size 128x16; Text 'HorizontalAlignment_2'
   Switch "HorizontalPictureAlignment" at 790,142 size 120x40; CaptionText 'Switch'; TextOff '0'; TextOn '1'
   TextField "Label_HorizontalPictureAlignment" at 790,184 size 128x16; Text 'HorizontalPictureAlignment'
   Switch "HorizontalPictureAlignment_2" at 920,142 size 120x40; CaptionText 'Switch'; TextOff '0'; TextOn '1'
   TextField "Label_HorizontalPictureAlignment_2" at 920,184 size 128x16; Text 'HorizontalPictureAlignment_2'
   Switch "InnerBackColorOff" at 1050,142 size 120x40; CaptionText 'Switch'; TextOff '0'; TextOn '1'
   TextField "Label_InnerBackColorOff" at 1050,184 size 128x16; Text 'InnerBackColorOff'
   Switch "InnerBackColorOn" at 10,208 size 120x40; CaptionText 'Switch'; TextOff '0'; TextOn '1'
   TextField "Label_InnerBackColorOn" at 10,250 size 128x16; Text 'InnerBackColorOn'
   Switch "MiddleGradientColor" at 140,208 size 120x40; CaptionText 'Switch'; TextOff '0'; TextOn '1'
   TextField "Label_MiddleGradientColor" at 140,250 size 128x16; Text 'MiddleGradientColor'
   Switch "PictureAreaBottomMargin" at 270,208 size 120x40; CaptionText 'Switch'; TextOff '0'; TextOn '1'
   TextField "Label_PictureAreaBottomMargin" at 270,250 size 128x16; Text 'PictureAreaBottomMargin'
   Switch "PictureAreaLeftMargin" at 400,208 size 120x40; CaptionText 'Switch'; TextOff '0'; TextOn '1'
   TextField "Label_PictureAreaLeftMargin" at 400,250 size 128x16; Text 'PictureAreaLeftMargin'
   Switch "PictureAreaRightMargin" at 530,208 size 120x40; CaptionText 'Switch'; TextOff '0'; TextOn '1'
   TextField "Label_PictureAreaRightMargin" at 530,250 size 128x16; Text 'PictureAreaRightMargin'
   Switch "PictureAreaTopMargin" at 660,208 size 120x40; CaptionText 'Switch'; TextOff '0'; TextOn '1'
   TextField "Label_PictureAreaTopMargin" at 660,250 size 128x16; Text 'PictureAreaTopMargin'
   Switch "SecondGradientColor" at 790,208 size 120x40; CaptionText 'Switch'; TextOff '0'; TextOn '1'
   TextField "Label_SecondGradientColor" at 790,250 size 128x16; Text 'SecondGradientColor'
   Switch "SecondGradientOffset" at 920,208 size 120x40; CaptionText 'Switch'; TextOff '0'; TextOn '1'
   TextField "Label_SecondGradientOffset" at 920,250 size 128x16; Text 'SecondGradientOffset'
   Switch "ShowCaption" at 1050,208 size 120x40; CaptionText 'Switch'; TextOff '0'; TextOn '1'
   TextField "Label_ShowCaption" at 1050,250 size 128x16; Text 'ShowCaption'
   Switch "SwitchOrientation" at 10,274 size 120x40; CaptionText 'Switch'; TextOff '0'; TextOn '1'
   TextField "Label_SwitchOrientation" at 10,316 size 128x16; Text 'SwitchOrientation'
   Switch "SwitchOrientation_2" at 140,274 size 120x40; CaptionText 'Switch'; TextOff '0'; TextOn '1'
   TextField "Label_SwitchOrientation_2" at 140,316 size 128x16; Text 'SwitchOrientation_2'
   Switch "SwitchOrientation_3" at 270,274 size 120x40; CaptionText 'Switch'; TextOff '0'; TextOn '1'
   TextField "Label_SwitchOrientation_3" at 270,316 size 128x16; Text 'SwitchOrientation_3'
   Switch "TextAreaBottomMargin" at 400,274 size 120x40; CaptionText 'Switch'; TextOff '0'; TextOn '1'
   TextField "Label_TextAreaBottomMargin" at 400,316 size 128x16; Text 'TextAreaBottomMargin'
   Switch "TextAreaLeftMargin" at 530,274 size 120x40; CaptionText 'Switch'; TextOff '0'; TextOn '1'
   TextField "Label_TextAreaLeftMargin" at 530,316 size 128x16; Text 'TextAreaLeftMargin'
   Switch "TextAreaRightMargin" at 660,274 size 120x40; CaptionText 'Switch'; TextOff '0'; TextOn '1'
   TextField "Label_TextAreaRightMargin" at 660,316 size 128x16; Text 'TextAreaRightMargin'
   Switch "TextAreaTopMargin" at 790,274 size 120x40; CaptionText 'Switch'; TextOff '0'; TextOn '1'
   TextField "Label_TextAreaTopMargin" at 790,316 size 128x16; Text 'TextAreaTopMargin'
   Switch "UseDesignColorSchema" at 920,274 size 120x40; CaptionText 'Switch'; TextOff '0'; TextOn '1'
   TextField "Label_UseDesignColorSchema" at 920,316 size 128x16; Text 'UseDesignColorSchema'
   Switch "UseFirstGradient" at 1050,274 size 120x40; CaptionText 'Switch'; TextOff '0'; TextOn '1'
   TextField "Label_UseFirstGradient" at 1050,316 size 128x16; Text 'UseFirstGradient'
   Switch "UseSecondGradient" at 10,340 size 120x40; CaptionText 'Switch'; TextOff '0'; TextOn '1'
   TextField "Label_UseSecondGradient" at 10,382 size 128x16; Text 'UseSecondGradient'
   Switch "VerticalAlignment" at 140,340 size 120x40; CaptionText 'Switch'; TextOff '0'; TextOn '1'
   TextField "Label_VerticalAlignment" at 140,382 size 128x16; Text 'VerticalAlignment'
   Switch "VerticalAlignment_2" at 270,340 size 120x40; CaptionText 'Switch'; TextOff '0'; TextOn '1'
   TextField "Label_VerticalAlignment_2" at 270,382 size 128x16; Text 'VerticalAlignment_2'
   Switch "VerticalPictureAlignment" at 400,340 size 120x40; CaptionText 'Switch'; TextOff '0'; TextOn '1'
   TextField "Label_VerticalPictureAlignment" at 400,382 size 128x16; Text 'VerticalPictureAlignment'
   Switch "VerticalPictureAlignment_2" at 530,340 size 120x40; CaptionText 'Switch'; TextOff '0'; TextOn '1'
   TextField "Label_VerticalPictureAlignment_2" at 530,382 size 128x16; Text 'VerticalPictureAlignment_2'
   Button "Next" at 1238,776 size 40x22; TextOff 'Text'
      on Click: ActivateScreen("P_SymbolLibrary_1", 0)

screen "P_SymbolLibrary_1" 1280x800
   SymbolLibrary "Default" at 10,10 size 60x60
   TextField "Label_Default" at 10,72 size 68x16; Text 'Default'
   SymbolLibrary "AboveUpperLimitColor" at 80,10 size 60x60
   TextField "Label_AboveUpperLimitColor" at 80,72 size 68x16; Text 'AboveUpperLimitColor'
   SymbolLibrary "BackColor" at 150,10 size 60x60
   TextField "Label_BackColor" at 150,72 size 68x16; Text 'BackColor'
   SymbolLibrary "BackFillStyle" at 220,10 size 60x60
   TextField "Label_BackFillStyle" at 220,72 size 68x16; Text 'BackFillStyle'
   SymbolLibrary "BelowLowerLimitColor" at 290,10 size 60x60
   TextField "Label_BelowLowerLimitColor" at 290,72 size 68x16; Text 'BelowLowerLimitColor'
   SymbolLibrary "BlinkColor" at 360,10 size 60x60
   TextField "Label_BlinkColor" at 360,72 size 68x16; Text 'BlinkColor'
   SymbolLibrary "FillColorMode" at 430,10 size 60x60
   TextField "Label_FillColorMode" at 430,72 size 68x16; Text 'FillColorMode'
   SymbolLibrary "FillColorMode_2" at 500,10 size 60x60
   TextField "Label_FillColorMode_2" at 500,72 size 68x16; Text 'FillColorMode_2'
   SymbolLibrary "FixedAspectRatio" at 570,10 size 60x60
   TextField "Label_FixedAspectRatio" at 570,72 size 68x16; Text 'FixedAspectRatio'
   SymbolLibrary "Flashing" at 640,10 size 60x60
   TextField "Label_Flashing" at 640,72 size 68x16; Text 'Flashing'
   SymbolLibrary "FlashingOnLimitViolation" at 710,10 size 60x60
   TextField "Label_FlashingOnLimitViolation" at 710,72 size 68x16; Text 'FlashingOnLimitViolation'
   SymbolLibrary "Flip" at 780,10 size 60x60
   TextField "Label_Flip" at 780,72 size 68x16; Text 'Flip'
   SymbolLibrary "Flip_2" at 850,10 size 60x60
   TextField "Label_Flip_2" at 850,72 size 68x16; Text 'Flip_2'
   SymbolLibrary "Flip_3" at 920,10 size 60x60
   TextField "Label_Flip_3" at 920,72 size 68x16; Text 'Flip_3'
   SymbolLibrary "ForeColor" at 990,10 size 60x60
   TextField "Label_ForeColor" at 990,72 size 68x16; Text 'ForeColor'
   SymbolLibrary "Rotation" at 1060,10 size 60x60
   TextField "Label_Rotation" at 1060,72 size 68x16; Text 'Rotation'
   SymbolLibrary "Rotation_2" at 1130,10 size 60x60
   TextField "Label_Rotation_2" at 1130,72 size 68x16; Text 'Rotation_2'
   SymbolLibrary "Rotation_3" at 1200,10 size 60x60
   TextField "Label_Rotation_3" at 1200,72 size 68x16; Text 'Rotation_3'
   Button "Next" at 1238,776 size 40x22; TextOff 'Text'
      on Click: ActivateScreen("P_Slider_1", 0)

screen "P_Slider_1" 1280x800
   Slider "Default" at 10,10 size 60x160; Caption 'SIMATIC'
   TextField "Label_Default" at 10,172 size 68x16; Text 'Default'
   Slider "BackColor" at 80,10 size 60x160; Caption 'SIMATIC'
   TextField "Label_BackColor" at 80,172 size 68x16; Text 'BackColor'
   Slider "BackFillStyle" at 150,10 size 60x160; Caption 'SIMATIC'
   TextField "Label_BackFillStyle" at 150,172 size 68x16; Text 'BackFillStyle'
   Slider "BarBackColor" at 220,10 size 60x160; Caption 'SIMATIC'
   TextField "Label_BarBackColor" at 220,172 size 68x16; Text 'BarBackColor'
   Slider "BarColor" at 290,10 size 60x160; Caption 'SIMATIC'
   TextField "Label_BarColor" at 290,172 size 68x16; Text 'BarColor'
   Slider "BarOrientation" at 360,10 size 60x160; Caption 'SIMATIC'
   TextField "Label_BarOrientation" at 360,172 size 68x16; Text 'BarOrientation'
   Slider "BarOrientation_2" at 430,10 size 60x160; Caption 'SIMATIC'
   TextField "Label_BarOrientation_2" at 430,172 size 68x16; Text 'BarOrientation_2'
   Slider "BarOrientation_3" at 500,10 size 60x160; Caption 'SIMATIC'
   TextField "Label_BarOrientation_3" at 500,172 size 68x16; Text 'BarOrientation_3'
   Slider "BorderBackColor" at 570,10 size 60x160; Caption 'SIMATIC'
   TextField "Label_BorderBackColor" at 570,172 size 68x16; Text 'BorderBackColor'
   Slider "BorderBrightColor3D" at 640,10 size 60x160; Caption 'SIMATIC'
   TextField "Label_BorderBrightColor3D" at 640,172 size 68x16; Text 'BorderBrightColor3D'
   Slider "BorderColor" at 710,10 size 60x160; Caption 'SIMATIC'
   TextField "Label_BorderColor" at 710,172 size 68x16; Text 'BorderColor'
   Slider "BorderInnerStyle3D" at 780,10 size 60x160; Caption 'SIMATIC'
   TextField "Label_BorderInnerStyle3D" at 780,172 size 68x16; Text 'BorderInnerStyle3D'
   Slider "BorderInnerStyle3D_2" at 850,10 size 60x160; Caption 'SIMATIC'
   TextField "Label_BorderInnerStyle3D_2" at 850,172 size 68x16; Text 'BorderInnerStyle3D_2'
   Slider "BorderInnerWidth3D" at 920,10 size 60x160; Caption 'SIMATIC'
   TextField "Label_BorderInnerWidth3D" at 920,172 size 68x16; Text 'BorderInnerWidth3D'
   Slider "BorderOuterStyle3D" at 990,10 size 60x160; Caption 'SIMATIC'
   TextField "Label_BorderOuterStyle3D" at 990,172 size 68x16; Text 'BorderOuterStyle3D'
   Slider "BorderOuterStyle3D_2" at 1060,10 size 60x160; Caption 'SIMATIC'
   TextField "Label_BorderOuterStyle3D_2" at 1060,172 size 68x16; Text 'BorderOuterStyle3D_2'
   Slider "BorderOuterWidth3D" at 1130,10 size 60x160; Caption 'SIMATIC'
   TextField "Label_BorderOuterWidth3D" at 1130,172 size 68x16; Text 'BorderOuterWidth3D'
   Slider "BorderShadeColor3D" at 1200,10 size 60x160; Caption 'SIMATIC'
   TextField "Label_BorderShadeColor3D" at 1200,172 size 68x16; Text 'BorderShadeColor3D'
   Slider "BorderWidth" at 10,196 size 60x160; Caption 'SIMATIC'
   TextField "Label_BorderWidth" at 10,358 size 68x16; Text 'BorderWidth'
   Slider "CornerRadius" at 80,196 size 60x160; Caption 'SIMATIC'
   TextField "Label_CornerRadius" at 80,358 size 68x16; Text 'CornerRadius'
   Slider "EdgeStyle" at 150,196 size 60x160; Caption 'SIMATIC'
   TextField "Label_EdgeStyle" at 150,358 size 68x16; Text 'EdgeStyle'
   Slider "EdgeStyle_2" at 220,196 size 60x160; Caption 'SIMATIC'
   TextField "Label_EdgeStyle_2" at 220,358 size 68x16; Text 'EdgeStyle_2'
   Slider "EdgeStyle_3" at 290,196 size 60x160; Caption 'SIMATIC'
   TextField "Label_EdgeStyle_3" at 290,358 size 68x16; Text 'EdgeStyle_3'
   Slider "EdgeStyle_4" at 360,196 size 60x160; Caption 'SIMATIC'
   TextField "Label_EdgeStyle_4" at 360,358 size 68x16; Text 'EdgeStyle_4'
   Slider "Flashing" at 430,196 size 60x160; Caption 'SIMATIC'
   TextField "Label_Flashing" at 430,358 size 68x16; Text 'Flashing'
   Slider "FocusColor" at 500,196 size 60x160; Caption 'SIMATIC'
   TextField "Label_FocusColor" at 500,358 size 68x16; Text 'FocusColor'
   Slider "FocusWidth" at 570,196 size 60x160; Caption 'SIMATIC'
   TextField "Label_FocusWidth" at 570,358 size 68x16; Text 'FocusWidth'
   Slider "ForeColor" at 640,196 size 60x160; Caption 'SIMATIC'
   TextField "Label_ForeColor" at 640,358 size 68x16; Text 'ForeColor'
   Slider "LabelColor" at 710,196 size 60x160; Caption 'SIMATIC'
   TextField "Label_LabelColor" at 710,358 size 68x16; Text 'LabelColor'
   Slider "MaximumValue" at 780,196 size 60x160; Caption 'SIMATIC'
   TextField "Label_MaximumValue" at 780,358 size 68x16; Text 'MaximumValue'
   Slider "MinimumValue" at 850,196 size 60x160; Caption 'SIMATIC'
   TextField "Label_MinimumValue" at 850,358 size 68x16; Text 'MinimumValue'
   Slider "RangeLower1Color" at 920,196 size 60x160; Caption 'SIMATIC'
   TextField "Label_RangeLower1Color" at 920,358 size 68x16; Text 'RangeLower1Color'
   Slider "RangeLower1Enabled" at 990,196 size 60x160; Caption 'SIMATIC'
   TextField "Label_RangeLower1Enabled" at 990,358 size 68x16; Text 'RangeLower1Enabled'
   Slider "RangeLower2Color" at 1060,196 size 60x160; Caption 'SIMATIC'
   TextField "Label_RangeLower2Color" at 1060,358 size 68x16; Text 'RangeLower2Color'
   Slider "RangeLower2Enabled" at 1130,196 size 60x160; Caption 'SIMATIC'
   TextField "Label_RangeLower2Enabled" at 1130,358 size 68x16; Text 'RangeLower2Enabled'
   Slider "RangeNormalColor" at 1200,196 size 60x160; Caption 'SIMATIC'
   TextField "Label_RangeNormalColor" at 1200,358 size 68x16; Text 'RangeNormalColor'
   Slider "RangeNormalEnabled" at 10,382 size 60x160; Caption 'SIMATIC'
   TextField "Label_RangeNormalEnabled" at 10,544 size 68x16; Text 'RangeNormalEnabled'
   Slider "RangeUpper1Color" at 80,382 size 60x160; Caption 'SIMATIC'
   TextField "Label_RangeUpper1Color" at 80,544 size 68x16; Text 'RangeUpper1Color'
   Slider "RangeUpper1Enabled" at 150,382 size 60x160; Caption 'SIMATIC'
   TextField "Label_RangeUpper1Enabled" at 150,544 size 68x16; Text 'RangeUpper1Enabled'
   Slider "RangeUpper2Color" at 220,382 size 60x160; Caption 'SIMATIC'
   TextField "Label_RangeUpper2Color" at 220,544 size 68x16; Text 'RangeUpper2Color'
   Slider "RangeUpper2Enabled" at 290,382 size 60x160; Caption 'SIMATIC'
   TextField "Label_RangeUpper2Enabled" at 290,544 size 68x16; Text 'RangeUpper2Enabled'
   Slider "ScalePosition" at 360,382 size 60x160; Caption 'SIMATIC'
   TextField "Label_ScalePosition" at 360,544 size 68x16; Text 'ScalePosition'
   Slider "ShowBar" at 430,382 size 60x160; Caption 'SIMATIC'
   TextField "Label_ShowBar" at 430,544 size 68x16; Text 'ShowBar'
   Slider "ShowLimitLines" at 500,382 size 60x160; Caption 'SIMATIC'
   TextField "Label_ShowLimitLines" at 500,544 size 68x16; Text 'ShowLimitLines'
   Slider "ShowLimitMarkers" at 570,382 size 60x160; Caption 'SIMATIC'
   TextField "Label_ShowLimitMarkers" at 570,544 size 68x16; Text 'ShowLimitMarkers'
   Slider "ShowLimitRanges" at 640,382 size 60x160; Caption 'SIMATIC'
   TextField "Label_ShowLimitRanges" at 640,544 size 68x16; Text 'ShowLimitRanges'
   Slider "ShowPosition" at 710,382 size 60x160; Caption 'SIMATIC'
   TextField "Label_ShowPosition" at 710,544 size 68x16; Text 'ShowPosition'
   Slider "ShowScale" at 780,382 size 60x160; Caption 'SIMATIC'
   TextField "Label_ShowScale" at 780,544 size 68x16; Text 'ShowScale'
   Slider "ShowThumb" at 850,382 size 60x160; Caption 'SIMATIC'
   TextField "Label_ShowThumb" at 850,544 size 68x16; Text 'ShowThumb'
   Slider "ShowTickLabels" at 920,382 size 60x160; Caption 'SIMATIC'
   TextField "Label_ShowTickLabels" at 920,544 size 68x16; Text 'ShowTickLabels'
   Slider "ShowTicks" at 990,382 size 60x160; Caption 'SIMATIC'
   TextField "Label_ShowTicks" at 990,544 size 68x16; Text 'ShowTicks'
   Slider "ThumbBackColor" at 1060,382 size 60x160; Caption 'SIMATIC'
   TextField "Label_ThumbBackColor" at 1060,544 size 68x16; Text 'ThumbBackColor'
   Slider "UseDesignColorSchema" at 1130,382 size 60x160; Caption 'SIMATIC'
   TextField "Label_UseDesignColorSchema" at 1130,544 size 68x16; Text 'UseDesignColorSchema'
   Button "Next" at 1238,776 size 40x22; TextOff 'Text'
      on Click: ActivateScreen("P_Gauge_1", 0)

screen "P_Gauge_1" 1280x800
   Gauge "Default" at 10,10 size 150x150; CaptionText 'SIMATIC'
   TextField "Label_Default" at 10,162 size 158x16; Text 'Default'
   Gauge "AngleMax" at 170,10 size 150x150; CaptionText 'SIMATIC'
   TextField "Label_AngleMax" at 170,162 size 158x16; Text 'AngleMax'
   Gauge "AngleMin" at 330,10 size 150x150; CaptionText 'SIMATIC'
   TextField "Label_AngleMin" at 330,162 size 158x16; Text 'AngleMin'
   Gauge "BackColor" at 490,10 size 150x150; CaptionText 'SIMATIC'
   TextField "Label_BackColor" at 490,162 size 158x16; Text 'BackColor'
   Gauge "BackFillStyle" at 650,10 size 150x150; CaptionText 'SIMATIC'
   TextField "Label_BackFillStyle" at 650,162 size 158x16; Text 'BackFillStyle'
   Gauge "BorderBackColor" at 810,10 size 150x150; CaptionText 'SIMATIC'
   TextField "Label_BorderBackColor" at 810,162 size 158x16; Text 'BorderBackColor'
   Gauge "BorderColor" at 970,10 size 150x150; CaptionText 'SIMATIC'
   TextField "Label_BorderColor" at 970,162 size 158x16; Text 'BorderColor'
   Gauge "BorderWidth" at 10,186 size 150x150; CaptionText 'SIMATIC'
   TextField "Label_BorderWidth" at 10,338 size 158x16; Text 'BorderWidth'
   Gauge "CaptionColor" at 170,186 size 150x150; CaptionText 'SIMATIC'
   TextField "Label_CaptionColor" at 170,338 size 158x16; Text 'CaptionColor'
   Gauge "CaptionTop" at 330,186 size 150x150; CaptionText 'SIMATIC'
   TextField "Label_CaptionTop" at 330,338 size 158x16; Text 'CaptionTop'
   Gauge "CenterColor" at 490,186 size 150x150; CaptionText 'SIMATIC'
   TextField "Label_CenterColor" at 490,338 size 158x16; Text 'CenterColor'
   Gauge "CenterSize" at 650,186 size 150x150; CaptionText 'SIMATIC'
   TextField "Label_CenterSize" at 650,338 size 158x16; Text 'CenterSize'
   Gauge "CornerRadius" at 810,186 size 150x150; CaptionText 'SIMATIC'
   TextField "Label_CornerRadius" at 810,338 size 158x16; Text 'CornerRadius'
   Gauge "DialColor" at 970,186 size 150x150; CaptionText 'SIMATIC'
   TextField "Label_DialColor" at 970,338 size 158x16; Text 'DialColor'
   Gauge "DialFillStyle" at 10,362 size 150x150; CaptionText 'SIMATIC'
   TextField "Label_DialFillStyle" at 10,514 size 158x16; Text 'DialFillStyle'
   Gauge "DialSize" at 170,362 size 150x150; CaptionText 'SIMATIC'
   TextField "Label_DialSize" at 170,514 size 158x16; Text 'DialSize'
   Gauge "EdgeStyle" at 330,362 size 150x150; CaptionText 'SIMATIC'
   TextField "Label_EdgeStyle" at 330,514 size 158x16; Text 'EdgeStyle'
   Gauge "EdgeStyle_2" at 490,362 size 150x150; CaptionText 'SIMATIC'
   TextField "Label_EdgeStyle_2" at 490,514 size 158x16; Text 'EdgeStyle_2'
   Gauge "EdgeStyle_3" at 650,362 size 150x150; CaptionText 'SIMATIC'
   TextField "Label_EdgeStyle_3" at 650,514 size 158x16; Text 'EdgeStyle_3'
   Gauge "EdgeStyle_4" at 810,362 size 150x150; CaptionText 'SIMATIC'
   TextField "Label_EdgeStyle_4" at 810,514 size 158x16; Text 'EdgeStyle_4'
   Gauge "Gradation" at 970,362 size 150x150; CaptionText 'SIMATIC'
   TextField "Label_Gradation" at 970,514 size 158x16; Text 'Gradation'
   Gauge "InnerDialColor" at 10,538 size 150x150; CaptionText 'SIMATIC'
   TextField "Label_InnerDialColor" at 10,690 size 158x16; Text 'InnerDialColor'
   Gauge "InnerDialInnerDistance" at 170,538 size 150x150; CaptionText 'SIMATIC'
   TextField "Label_InnerDialInnerDistance" at 170,690 size 158x16; Text 'InnerDialInnerDistance'
   Gauge "InnerDialOuterDistance" at 330,538 size 150x150; CaptionText 'SIMATIC'
   TextField "Label_InnerDialOuterDistance" at 330,690 size 158x16; Text 'InnerDialOuterDistance'
   Gauge "LockSquaredExtent" at 490,538 size 150x150; CaptionText 'SIMATIC'
   TextField "Label_LockSquaredExtent" at 490,690 size 158x16; Text 'LockSquaredExtent'
   Gauge "MaximumValue" at 650,538 size 150x150; CaptionText 'SIMATIC'
   TextField "Label_MaximumValue" at 650,690 size 158x16; Text 'MaximumValue'
   Gauge "MinimumValue" at 810,538 size 150x150; CaptionText 'SIMATIC'
   TextField "Label_MinimumValue" at 810,690 size 158x16; Text 'MinimumValue'
   Gauge "NeedleHeight" at 970,538 size 150x150; CaptionText 'SIMATIC'
   TextField "Label_NeedleHeight" at 970,690 size 158x16; Text 'NeedleHeight'
   Button "Next" at 1238,776 size 40x22; TextOff 'Text'
      on Click: ActivateScreen("P_Gauge_2", 0)

screen "P_Gauge_2" 1280x800
   Gauge "PointerColor" at 10,10 size 150x150; CaptionText 'SIMATIC'
   TextField "Label_PointerColor" at 10,162 size 158x16; Text 'PointerColor'
   Gauge "RangeLower1Color" at 170,10 size 150x150; CaptionText 'SIMATIC'
   TextField "Label_RangeLower1Color" at 170,162 size 158x16; Text 'RangeLower1Color'
   Gauge "RangeLower1Enabled" at 330,10 size 150x150; CaptionText 'SIMATIC'
   TextField "Label_RangeLower1Enabled" at 330,162 size 158x16; Text 'RangeLower1Enabled'
   Gauge "RangeLower2Color" at 490,10 size 150x150; CaptionText 'SIMATIC'
   TextField "Label_RangeLower2Color" at 490,162 size 158x16; Text 'RangeLower2Color'
   Gauge "RangeLower2Enabled" at 650,10 size 150x150; CaptionText 'SIMATIC'
   TextField "Label_RangeLower2Enabled" at 650,162 size 158x16; Text 'RangeLower2Enabled'
   Gauge "RangeNormalColor" at 810,10 size 150x150; CaptionText 'SIMATIC'
   TextField "Label_RangeNormalColor" at 810,162 size 158x16; Text 'RangeNormalColor'
   Gauge "RangeNormalEnabled" at 970,10 size 150x150; CaptionText 'SIMATIC'
   TextField "Label_RangeNormalEnabled" at 970,162 size 158x16; Text 'RangeNormalEnabled'
   Gauge "RangeUpper1Color" at 10,186 size 150x150; CaptionText 'SIMATIC'
   TextField "Label_RangeUpper1Color" at 10,338 size 158x16; Text 'RangeUpper1Color'
   Gauge "RangeUpper1Enabled" at 170,186 size 150x150; CaptionText 'SIMATIC'
   TextField "Label_RangeUpper1Enabled" at 170,338 size 158x16; Text 'RangeUpper1Enabled'
   Gauge "RangeUpper1Start" at 330,186 size 150x150; CaptionText 'SIMATIC'
   TextField "Label_RangeUpper1Start" at 330,338 size 158x16; Text 'RangeUpper1Start'
   Gauge "RangeUpper2Color" at 490,186 size 150x150; CaptionText 'SIMATIC'
   TextField "Label_RangeUpper2Color" at 490,338 size 158x16; Text 'RangeUpper2Color'
   Gauge "RangeUpper2Enabled" at 650,186 size 150x150; CaptionText 'SIMATIC'
   TextField "Label_RangeUpper2Enabled" at 650,338 size 158x16; Text 'RangeUpper2Enabled'
   Gauge "RangeUpper2Start" at 810,186 size 150x150; CaptionText 'SIMATIC'
   TextField "Label_RangeUpper2Start" at 810,338 size 158x16; Text 'RangeUpper2Start'
   Gauge "ScaleLabelColor" at 970,186 size 150x150; CaptionText 'SIMATIC'
   TextField "Label_ScaleLabelColor" at 970,338 size 158x16; Text 'ScaleLabelColor'
   Gauge "ScaleTickColor" at 10,362 size 150x150; CaptionText 'SIMATIC'
   TextField "Label_ScaleTickColor" at 10,514 size 158x16; Text 'ScaleTickColor'
   Gauge "ScaleTickLabelPosition" at 170,362 size 150x150; CaptionText 'SIMATIC'
   TextField "Label_ScaleTickLabelPosition" at 170,514 size 158x16; Text 'ScaleTickLabelPosition'
   Gauge "ScaleTickLength" at 330,362 size 150x150; CaptionText 'SIMATIC'
   TextField "Label_ScaleTickLength" at 330,514 size 158x16; Text 'ScaleTickLength'
   Gauge "ScaleTickPosition" at 490,362 size 150x150; CaptionText 'SIMATIC'
   TextField "Label_ScaleTickPosition" at 490,514 size 158x16; Text 'ScaleTickPosition'
   Gauge "ShowDecimalPoint" at 650,362 size 150x150; CaptionText 'SIMATIC'
   TextField "Label_ShowDecimalPoint" at 650,514 size 158x16; Text 'ShowDecimalPoint'
   Gauge "ShowInnerDial" at 810,362 size 150x150; CaptionText 'SIMATIC'
   TextField "Label_ShowInnerDial" at 810,514 size 158x16; Text 'ShowInnerDial'
   Gauge "ShowLimitRanges" at 970,362 size 150x150; CaptionText 'SIMATIC'
   TextField "Label_ShowLimitRanges" at 970,514 size 158x16; Text 'ShowLimitRanges'
   Gauge "ShowPeakValuePointer" at 10,538 size 150x150; CaptionText 'SIMATIC'
   TextField "Label_ShowPeakValuePointer" at 10,690 size 158x16; Text 'ShowPeakValuePointer'
   Gauge "UnitColor" at 170,538 size 150x150; CaptionText 'SIMATIC'
   TextField "Label_UnitColor" at 170,690 size 158x16; Text 'UnitColor'
   Gauge "UnitTop" at 330,538 size 150x150; CaptionText 'SIMATIC'
   TextField "Label_UnitTop" at 330,690 size 158x16; Text 'UnitTop'
   Gauge "UseDesignColorSchema" at 490,538 size 150x150; CaptionText 'SIMATIC'
   TextField "Label_UseDesignColorSchema" at 490,690 size 158x16; Text 'UseDesignColorSchema'
   Button "Next" at 1238,776 size 40x22; TextOff 'Text'
      on Click: ActivateScreen("P_Clock_1", 0)

screen "P_Clock_1" 1280x800
   Clock "Default" at 10,10 size 150x150
   TextField "Label_Default" at 10,162 size 158x16; Text 'Default'
   Clock "Analog" at 170,10 size 150x150
   TextField "Label_Analog" at 170,162 size 158x16; Text 'Analog'
   Clock "BackFillStyle" at 330,10 size 150x150
   TextField "Label_BackFillStyle" at 330,162 size 158x16; Text 'BackFillStyle'
   Clock "BorderBackColor" at 490,10 size 150x150
   TextField "Label_BorderBackColor" at 490,162 size 158x16; Text 'BorderBackColor'
   Clock "BorderColor" at 650,10 size 150x150
   TextField "Label_BorderColor" at 650,162 size 158x16; Text 'BorderColor'
   Clock "BorderWidth" at 810,10 size 150x150
   TextField "Label_BorderWidth" at 810,162 size 158x16; Text 'BorderWidth'
   Clock "CornerRadius" at 970,10 size 150x150
   TextField "Label_CornerRadius" at 970,162 size 158x16; Text 'CornerRadius'
   Clock "DialColor" at 10,186 size 150x150
   TextField "Label_DialColor" at 10,338 size 158x16; Text 'DialColor'
   Clock "EdgeStyle" at 170,186 size 150x150
   TextField "Label_EdgeStyle" at 170,338 size 158x16; Text 'EdgeStyle'
   Clock "EdgeStyle_2" at 330,186 size 150x150
   TextField "Label_EdgeStyle_2" at 330,338 size 158x16; Text 'EdgeStyle_2'
   Clock "EdgeStyle_3" at 490,186 size 150x150
   TextField "Label_EdgeStyle_3" at 490,338 size 158x16; Text 'EdgeStyle_3'
   Clock "EdgeStyle_4" at 650,186 size 150x150
   TextField "Label_EdgeStyle_4" at 650,338 size 158x16; Text 'EdgeStyle_4'
   Clock "Flashing" at 810,186 size 150x150
   TextField "Label_Flashing" at 810,338 size 158x16; Text 'Flashing'
   Clock "HourNeedleHeight" at 970,186 size 150x150
   TextField "Label_HourNeedleHeight" at 970,338 size 158x16; Text 'HourNeedleHeight'
   Clock "HourNeedleWidth" at 10,362 size 150x150
   TextField "Label_HourNeedleWidth" at 10,514 size 158x16; Text 'HourNeedleWidth'
   Clock "LockSquaredExtent" at 170,362 size 150x150
   TextField "Label_LockSquaredExtent" at 170,514 size 158x16; Text 'LockSquaredExtent'
   Clock "MinuteNeedleHeight" at 330,362 size 150x150
   TextField "Label_MinuteNeedleHeight" at 330,514 size 158x16; Text 'MinuteNeedleHeight'
   Clock "MinuteNeedleWidth" at 490,362 size 150x150
   TextField "Label_MinuteNeedleWidth" at 490,514 size 158x16; Text 'MinuteNeedleWidth'
   Clock "NeedleBorderColor" at 650,362 size 150x150
   TextField "Label_NeedleBorderColor" at 650,514 size 158x16; Text 'NeedleBorderColor'
   Clock "NeedleColor" at 810,362 size 150x150
   TextField "Label_NeedleColor" at 810,514 size 158x16; Text 'NeedleColor'
   Clock "NeedleFillStyle" at 970,362 size 150x150
   TextField "Label_NeedleFillStyle" at 970,514 size 158x16; Text 'NeedleFillStyle'
   Clock "NumberStyle" at 10,538 size 150x150
   TextField "Label_NumberStyle" at 10,690 size 158x16; Text 'NumberStyle'
   Clock "NumberStyle_2" at 170,538 size 150x150
   TextField "Label_NumberStyle_2" at 170,690 size 158x16; Text 'NumberStyle_2'
   Clock "SecondNeedleHeight" at 330,538 size 150x150
   TextField "Label_SecondNeedleHeight" at 330,690 size 158x16; Text 'SecondNeedleHeight'
   Clock "SecondNeedleWidth" at 490,538 size 150x150
   TextField "Label_SecondNeedleWidth" at 490,690 size 158x16; Text 'SecondNeedleWidth'
   Clock "ShowTicks" at 650,538 size 150x150
   TextField "Label_ShowTicks" at 650,690 size 158x16; Text 'ShowTicks'
   Clock "TickDistance" at 810,538 size 150x150
   TextField "Label_TickDistance" at 810,690 size 158x16; Text 'TickDistance'
   Clock "TickStyle" at 970,538 size 150x150
   TextField "Label_TickStyle" at 970,690 size 158x16; Text 'TickStyle'
   Button "Next" at 1238,776 size 40x22; TextOff 'Text'
      on Click: ActivateScreen("P_Clock_2", 0)

screen "P_Clock_2" 1280x800
   Clock "TicksColor" at 10,10 size 150x150
   TextField "Label_TicksColor" at 10,162 size 158x16; Text 'TicksColor'
   Clock "UseDesignColorSchema" at 170,10 size 150x150
   TextField "Label_UseDesignColorSchema" at 170,162 size 158x16; Text 'UseDesignColorSchema'
   Button "Next" at 1238,776 size 40x22; TextOff 'Text'
      on Click: ActivateScreen("P_Line_1", 0)

screen "D_Bar_1" 1280x800
   Bar "Static" at 6,4 size 40x120
   TextField "Label_Static" at 6,156 size 88x16; Text 'Static'
   Bar "A_Range" at 98,4 size 40x120
      Appearance <- "D_Range"
   TextField "Label_A_Range" at 98,156 size 88x16; Text 'A_Range'
   Bar "A_Flash" at 190,4 size 40x120
      Appearance <- "D_Range"
   TextField "Label_A_Flash" at 190,156 size 88x16; Text 'A_Flash'
   Bar "A_Bit" at 282,4 size 40x120
      Appearance <- "D_Bool"
   TextField "Label_A_Bit" at 282,156 size 88x16; Text 'A_Bit'
   Bar "A_Bits" at 374,4 size 40x120
      Appearance <- "D_Bits"
   TextField "Label_A_Bits" at 374,156 size 88x16; Text 'A_Bits'
   Bar "V_Range" at 466,4 size 40x120
      Visibility <- "D_Range"
   TextField "Label_V_Range" at 466,156 size 88x16; Text 'V_Range'
   Bar "V_Bit" at 558,4 size 40x120
      Visibility <- "D_Vis"
   TextField "Label_V_Bit" at 558,156 size 88x16; Text 'V_Bit'
   Bar "M_H" at 650,4 size 40x120
      HorizontalMovement <- "D_Pct"
   TextField "Label_M_H" at 650,156 size 88x16; Text 'M_H'
   Bar "M_V" at 742,4 size 40x120
      VerticalMovement <- "D_Pct"
   TextField "Label_M_V" at 742,156 size 88x16; Text 'M_V'
   Bar "M_D" at 834,4 size 40x120
      DiagonalMovement <- "D_Pct"
   TextField "Label_M_D" at 834,156 size 88x16; Text 'M_D'
   Bar "M_Direct" at 926,4 size 40x120
      DirectMovement <- "D_X"
      DirectMovement <- "D_Y"
   TextField "Label_M_Direct" at 926,156 size 88x16; Text 'M_Direct'
   Bar "E_Range" at 1018,4 size 40x120
      ObjectEnable <- "D_Range"
   TextField "Label_E_Range" at 1018,156 size 88x16; Text 'E_Range'
   Bar "E_Bit" at 1110,4 size 40x120
      ObjectEnable <- "D_En"
   TextField "Label_E_Bit" at 1110,156 size 88x16; Text 'E_Bit'
   Bar "PV_Pct" at 6,176 size 40x120
      ProcessValue <- "D_Pct"
   TextField "Label_PV_Pct" at 6,328 size 88x16; Text 'PV_Pct'
   Bar "PV_Real" at 98,176 size 40x120
      ProcessValue <- "D_Real"
   TextField "Label_PV_Real" at 98,328 size 88x16; Text 'PV_Real'
   Bar "PV_BarR" at 190,176 size 40x120
      ProcessValue <- "D_BarR"
   TextField "Label_PV_BarR" at 190,328 size 88x16; Text 'PV_BarR'
   Bar "PV_Pct_0_100" at 282,176 size 40x120; MinimumValue 0; MaximumValue 100
      ProcessValue <- "D_Pct"
   TextField "Label_PV_Pct_0_100" at 282,328 size 88x16; Text 'PV_Pct_0_100'
   Bar "PV_Pct_MaxMin" at 374,176 size 40x120
      ProcessValue <- "D_Pct"
      MaximumValue <- "D_Max"
      MinimumValue <- "D_Min"
   TextField "Label_PV_Pct_MaxMin" at 374,328 size 88x16; Text 'PV_Pct_MaxMin'
   IOField "State" at 4,774 size 60x22; FormatPattern 9
      ProcessValue <- "D_State"
   Button "S1" at 70,774 size 40x22; TextOff 'S1'
      on Click: "SetS1"()
   Button "S2" at 114,774 size 40x22; TextOff 'S2'
      on Click: "SetS2"()
   Button "S3" at 158,774 size 40x22; TextOff 'S3'
      on Click: "SetS3"()
   Button "S4" at 202,774 size 40x22; TextOff 'S4'
      on Click: "SetS4"()
   Button "Next" at 1236,774 size 40x22; TextOff 'Next'
      on Click: ActivateScreen("D_Switch_1", 0)

screen "D_Button_1" 1280x800
   Button "Static" at 6,4 size 100x40; TextOff 'Text'
   TextField "Label_Static" at 6,76 size 148x16; Text 'Static'
   Button "A_Range" at 158,4 size 100x40; TextOff 'Text'
      Appearance <- "D_Range"
   TextField "Label_A_Range" at 158,76 size 148x16; Text 'A_Range'
   Button "A_Flash" at 310,4 size 100x40; TextOff 'Text'
      Appearance <- "D_Range"
   TextField "Label_A_Flash" at 310,76 size 148x16; Text 'A_Flash'
   Button "A_Bit" at 462,4 size 100x40; TextOff 'Text'
      Appearance <- "D_Bool"
   TextField "Label_A_Bit" at 462,76 size 148x16; Text 'A_Bit'
   Button "A_Bits" at 614,4 size 100x40; TextOff 'Text'
      Appearance <- "D_Bits"
   TextField "Label_A_Bits" at 614,76 size 148x16; Text 'A_Bits'
   Button "V_Range" at 766,4 size 100x40; TextOff 'Text'
      Visibility <- "D_Range"
   TextField "Label_V_Range" at 766,76 size 148x16; Text 'V_Range'
   Button "V_Bit" at 918,4 size 100x40; TextOff 'Text'
      Visibility <- "D_Vis"
   TextField "Label_V_Bit" at 918,76 size 148x16; Text 'V_Bit'
   Button "M_H" at 1070,4 size 100x40; TextOff 'Text'
      HorizontalMovement <- "D_Pct"
   TextField "Label_M_H" at 1070,76 size 148x16; Text 'M_H'
   Button "M_V" at 6,96 size 100x40; TextOff 'Text'
      VerticalMovement <- "D_Pct"
   TextField "Label_M_V" at 6,168 size 148x16; Text 'M_V'
   Button "M_D" at 158,96 size 100x40; TextOff 'Text'
      DiagonalMovement <- "D_Pct"
   TextField "Label_M_D" at 158,168 size 148x16; Text 'M_D'
   Button "M_Direct" at 310,96 size 100x40; TextOff 'Text'
      DirectMovement <- "D_X"
      DirectMovement <- "D_Y"
   TextField "Label_M_Direct" at 310,168 size 148x16; Text 'M_Direct'
   Button "E_Range" at 462,96 size 100x40; TextOff 'Text'
      ObjectEnable <- "D_Range"
   TextField "Label_E_Range" at 462,168 size 148x16; Text 'E_Range'
   Button "E_Bit" at 614,96 size 100x40; TextOff 'Text'
      ObjectEnable <- "D_En"
   TextField "Label_E_Bit" at 614,168 size 148x16; Text 'E_Bit'
   IOField "State" at 4,774 size 60x22; FormatPattern 9
      ProcessValue <- "D_State"
   Button "S1" at 70,774 size 40x22; TextOff 'S1'
      on Click: "SetS1"()
   Button "S2" at 114,774 size 40x22; TextOff 'S2'
      on Click: "SetS2"()
   Button "S3" at 158,774 size 40x22; TextOff 'S3'
      on Click: "SetS3"()
   Button "S4" at 202,774 size 40x22; TextOff 'S4'
      on Click: "SetS4"()
   Button "Next" at 1236,774 size 40x22; TextOff 'Next'
      on Click: ActivateScreen("D_SymbolicIOField_1", 0)

screen "D_Circle_1" 1280x800
   TextField "Label_Static" at 6,86 size 98x16; Text 'Static'
   Circle "A_Range" at 108,4 size 50x50
      Appearance <- "D_Range"
   TextField "Label_A_Range" at 108,86 size 98x16; Text 'A_Range'
   Circle "A_Flash" at 210,4 size 50x50
      Appearance <- "D_Range"
   TextField "Label_A_Flash" at 210,86 size 98x16; Text 'A_Flash'
   Circle "A_Bit" at 312,4 size 50x50
      Appearance <- "D_Bool"
   TextField "Label_A_Bit" at 312,86 size 98x16; Text 'A_Bit'
   Circle "A_Bits" at 414,4 size 50x50
      Appearance <- "D_Bits"
   TextField "Label_A_Bits" at 414,86 size 98x16; Text 'A_Bits'
   Circle "V_Range" at 516,4 size 50x50
      Visibility <- "D_Range"
   TextField "Label_V_Range" at 516,86 size 98x16; Text 'V_Range'
   Circle "V_Bit" at 618,4 size 50x50
      Visibility <- "D_Vis"
   TextField "Label_V_Bit" at 618,86 size 98x16; Text 'V_Bit'
   Circle "M_H" at 720,4 size 50x50
      HorizontalMovement <- "D_Pct"
   TextField "Label_M_H" at 720,86 size 98x16; Text 'M_H'
   Circle "M_V" at 822,4 size 50x50
      VerticalMovement <- "D_Pct"
   TextField "Label_M_V" at 822,86 size 98x16; Text 'M_V'
   Circle "M_D" at 924,4 size 50x50
      DiagonalMovement <- "D_Pct"
   TextField "Label_M_D" at 924,86 size 98x16; Text 'M_D'
   Circle "M_Direct" at 1026,4 size 50x50
      DirectMovement <- "D_X"
      DirectMovement <- "D_Y"
   TextField "Label_M_Direct" at 1026,86 size 98x16; Text 'M_Direct'
   Circle "E_Range" at 1128,4 size 50x50
      ObjectEnable <- "D_Range"
   TextField "Label_E_Range" at 1128,86 size 98x16; Text 'E_Range'
   Circle "E_Bit" at 6,106 size 50x50
      ObjectEnable <- "D_En"
   TextField "Label_E_Bit" at 6,188 size 98x16; Text 'E_Bit'
   IOField "State" at 4,774 size 60x22; FormatPattern 9
      ProcessValue <- "D_State"
   Button "S1" at 70,774 size 40x22; TextOff 'S1'
      on Click: "SetS1"()
   Button "S2" at 114,774 size 40x22; TextOff 'S2'
      on Click: "SetS2"()
   Button "S3" at 158,774 size 40x22; TextOff 'S3'
      on Click: "SetS3"()
   Button "S4" at 202,774 size 40x22; TextOff 'S4'
      on Click: "SetS4"()
   Button "Next" at 1236,774 size 40x22; TextOff 'Next'
      on Click: ActivateScreen("D_Rectangle_1", 0)

screen "D_Clock_1" 1280x800
   Clock "Static" at 6,4 size 150x150
   TextField "Label_Static" at 6,186 size 198x16; Text 'Static'
   Clock "A_Range" at 208,4 size 150x150
      Appearance <- "D_Range"
   TextField "Label_A_Range" at 208,186 size 198x16; Text 'A_Range'
   Clock "A_Flash" at 410,4 size 150x150
      Appearance <- "D_Range"
   TextField "Label_A_Flash" at 410,186 size 198x16; Text 'A_Flash'
   Clock "A_Bit" at 612,4 size 150x150
      Appearance <- "D_Bool"
   TextField "Label_A_Bit" at 612,186 size 198x16; Text 'A_Bit'
   Clock "A_Bits" at 814,4 size 150x150
      Appearance <- "D_Bits"
   TextField "Label_A_Bits" at 814,186 size 198x16; Text 'A_Bits'
   Clock "V_Range" at 1016,4 size 150x150
      Visibility <- "D_Range"
   TextField "Label_V_Range" at 1016,186 size 198x16; Text 'V_Range'
   Clock "V_Bit" at 6,206 size 150x150
      Visibility <- "D_Vis"
   TextField "Label_V_Bit" at 6,388 size 198x16; Text 'V_Bit'
   Clock "M_H" at 208,206 size 150x150
      HorizontalMovement <- "D_Pct"
   TextField "Label_M_H" at 208,388 size 198x16; Text 'M_H'
   Clock "M_V" at 410,206 size 150x150
      VerticalMovement <- "D_Pct"
   TextField "Label_M_V" at 410,388 size 198x16; Text 'M_V'
   Clock "M_D" at 612,206 size 150x150
      DiagonalMovement <- "D_Pct"
   TextField "Label_M_D" at 612,388 size 198x16; Text 'M_D'
   Clock "M_Direct" at 814,206 size 150x150
      DirectMovement <- "D_X"
      DirectMovement <- "D_Y"
   TextField "Label_M_Direct" at 814,388 size 198x16; Text 'M_Direct'
   Clock "E_Range" at 1016,206 size 150x150
      ObjectEnable <- "D_Range"
   TextField "Label_E_Range" at 1016,388 size 198x16; Text 'E_Range'
   Clock "E_Bit" at 6,408 size 150x150
      ObjectEnable <- "D_En"
   TextField "Label_E_Bit" at 6,590 size 198x16; Text 'E_Bit'
   IOField "State" at 4,774 size 60x22; FormatPattern 9
      ProcessValue <- "D_State"
   Button "S1" at 70,774 size 40x22; TextOff 'S1'
      on Click: "SetS1"()
   Button "S2" at 114,774 size 40x22; TextOff 'S2'
      on Click: "SetS2"()
   Button "S3" at 158,774 size 40x22; TextOff 'S3'
      on Click: "SetS3"()
   Button "S4" at 202,774 size 40x22; TextOff 'S4'
      on Click: "SetS4"()
   Button "Next" at 1236,774 size 40x22; TextOff 'Next'
      on Click: ActivateScreen("D_Line_1", 0)

screen "D_DateTimeField_1" 1280x800
   DateTimeField "Static" at 6,4 size 160x30
   TextField "Label_Static" at 6,66 size 208x16; Text 'Static'
   DateTimeField "A_Range" at 218,4 size 160x30
      Appearance <- "D_Range"
   TextField "Label_A_Range" at 218,66 size 208x16; Text 'A_Range'
   DateTimeField "A_Flash" at 430,4 size 160x30
      Appearance <- "D_Range"
   TextField "Label_A_Flash" at 430,66 size 208x16; Text 'A_Flash'
   DateTimeField "A_Bit" at 642,4 size 160x30
      Appearance <- "D_Bool"
   TextField "Label_A_Bit" at 642,66 size 208x16; Text 'A_Bit'
   DateTimeField "A_Bits" at 854,4 size 160x30
      Appearance <- "D_Bits"
   TextField "Label_A_Bits" at 854,66 size 208x16; Text 'A_Bits'
   DateTimeField "V_Range" at 1066,4 size 160x30
      Visibility <- "D_Range"
   TextField "Label_V_Range" at 1066,66 size 208x16; Text 'V_Range'
   DateTimeField "V_Bit" at 6,86 size 160x30
      Visibility <- "D_Vis"
   TextField "Label_V_Bit" at 6,148 size 208x16; Text 'V_Bit'
   DateTimeField "M_H" at 218,86 size 160x30
      HorizontalMovement <- "D_Pct"
   TextField "Label_M_H" at 218,148 size 208x16; Text 'M_H'
   DateTimeField "M_V" at 430,86 size 160x30
      VerticalMovement <- "D_Pct"
   TextField "Label_M_V" at 430,148 size 208x16; Text 'M_V'
   DateTimeField "M_D" at 642,86 size 160x30
      DiagonalMovement <- "D_Pct"
   TextField "Label_M_D" at 642,148 size 208x16; Text 'M_D'
   DateTimeField "M_Direct" at 854,86 size 160x30
      DirectMovement <- "D_X"
      DirectMovement <- "D_Y"
   TextField "Label_M_Direct" at 854,148 size 208x16; Text 'M_Direct'
   DateTimeField "E_Range" at 1066,86 size 160x30
      ObjectEnable <- "D_Range"
   TextField "Label_E_Range" at 1066,148 size 208x16; Text 'E_Range'
   DateTimeField "E_Bit" at 6,168 size 160x30
      ObjectEnable <- "D_En"
   TextField "Label_E_Bit" at 6,230 size 208x16; Text 'E_Bit'
   DateTimeField "PV_DateTime" at 218,168 size 160x30
      ProcessValue <- "D_DateTime"
   TextField "Label_PV_DateTime" at 218,230 size 208x16; Text 'PV_DateTime'
   IOField "State" at 4,774 size 60x22; FormatPattern 9
      ProcessValue <- "D_State"
   Button "S1" at 70,774 size 40x22; TextOff 'S1'
      on Click: "SetS1"()
   Button "S2" at 114,774 size 40x22; TextOff 'S2'
      on Click: "SetS2"()
   Button "S3" at 158,774 size 40x22; TextOff 'S3'
      on Click: "SetS3"()
   Button "S4" at 202,774 size 40x22; TextOff 'S4'
      on Click: "SetS4"()
   Button "Next" at 1236,774 size 40x22; TextOff 'Next'
      on Click: ActivateScreen("D_Bar_1", 0)

screen "D_Ellipse_1" 1280x800
   TextField "Label_Static" at 6,86 size 148x16; Text 'Static'
   Ellipse "A_Range" at 158,4 size 100x50
      Appearance <- "D_Range"
   TextField "Label_A_Range" at 158,86 size 148x16; Text 'A_Range'
   Ellipse "A_Flash" at 310,4 size 100x50
      Appearance <- "D_Range"
   TextField "Label_A_Flash" at 310,86 size 148x16; Text 'A_Flash'
   Ellipse "A_Bit" at 462,4 size 100x50
      Appearance <- "D_Bool"
   TextField "Label_A_Bit" at 462,86 size 148x16; Text 'A_Bit'
   Ellipse "A_Bits" at 614,4 size 100x50
      Appearance <- "D_Bits"
   TextField "Label_A_Bits" at 614,86 size 148x16; Text 'A_Bits'
   Ellipse "V_Range" at 766,4 size 100x50
      Visibility <- "D_Range"
   TextField "Label_V_Range" at 766,86 size 148x16; Text 'V_Range'
   Ellipse "V_Bit" at 918,4 size 100x50
      Visibility <- "D_Vis"
   TextField "Label_V_Bit" at 918,86 size 148x16; Text 'V_Bit'
   Ellipse "M_H" at 1070,4 size 100x50
      HorizontalMovement <- "D_Pct"
   TextField "Label_M_H" at 1070,86 size 148x16; Text 'M_H'
   Ellipse "M_V" at 6,106 size 100x50
      VerticalMovement <- "D_Pct"
   TextField "Label_M_V" at 6,188 size 148x16; Text 'M_V'
   Ellipse "M_D" at 158,106 size 100x50
      DiagonalMovement <- "D_Pct"
   TextField "Label_M_D" at 158,188 size 148x16; Text 'M_D'
   Ellipse "M_Direct" at 310,106 size 100x50
      DirectMovement <- "D_X"
      DirectMovement <- "D_Y"
   TextField "Label_M_Direct" at 310,188 size 148x16; Text 'M_Direct'
   Ellipse "E_Range" at 462,106 size 100x50
      ObjectEnable <- "D_Range"
   TextField "Label_E_Range" at 462,188 size 148x16; Text 'E_Range'
   Ellipse "E_Bit" at 614,106 size 100x50
      ObjectEnable <- "D_En"
   TextField "Label_E_Bit" at 614,188 size 148x16; Text 'E_Bit'
   IOField "State" at 4,774 size 60x22; FormatPattern 9
      ProcessValue <- "D_State"
   Button "S1" at 70,774 size 40x22; TextOff 'S1'
      on Click: "SetS1"()
   Button "S2" at 114,774 size 40x22; TextOff 'S2'
      on Click: "SetS2"()
   Button "S3" at 158,774 size 40x22; TextOff 'S3'
      on Click: "SetS3"()
   Button "S4" at 202,774 size 40x22; TextOff 'S4'
      on Click: "SetS4"()
   Button "Next" at 1236,774 size 40x22; TextOff 'Next'
      on Click: ActivateScreen("D_Circle_1", 0)

screen "D_Gauge_1" 1280x800
   Gauge "Static" at 6,4 size 150x150; CaptionText 'SIMATIC'
   TextField "Label_Static" at 6,186 size 198x16; Text 'Static'
   Gauge "A_Range" at 208,4 size 150x150; CaptionText 'SIMATIC'
      Appearance <- "D_Range"
   TextField "Label_A_Range" at 208,186 size 198x16; Text 'A_Range'
   Gauge "A_Flash" at 410,4 size 150x150; CaptionText 'SIMATIC'
      Appearance <- "D_Range"
   TextField "Label_A_Flash" at 410,186 size 198x16; Text 'A_Flash'
   Gauge "A_Bit" at 612,4 size 150x150; CaptionText 'SIMATIC'
      Appearance <- "D_Bool"
   TextField "Label_A_Bit" at 612,186 size 198x16; Text 'A_Bit'
   Gauge "A_Bits" at 814,4 size 150x150; CaptionText 'SIMATIC'
      Appearance <- "D_Bits"
   TextField "Label_A_Bits" at 814,186 size 198x16; Text 'A_Bits'
   Gauge "V_Range" at 1016,4 size 150x150; CaptionText 'SIMATIC'
      Visibility <- "D_Range"
   TextField "Label_V_Range" at 1016,186 size 198x16; Text 'V_Range'
   Gauge "V_Bit" at 6,206 size 150x150; CaptionText 'SIMATIC'
      Visibility <- "D_Vis"
   TextField "Label_V_Bit" at 6,388 size 198x16; Text 'V_Bit'
   Gauge "M_H" at 208,206 size 150x150; CaptionText 'SIMATIC'
      HorizontalMovement <- "D_Pct"
   TextField "Label_M_H" at 208,388 size 198x16; Text 'M_H'
   Gauge "M_V" at 410,206 size 150x150; CaptionText 'SIMATIC'
      VerticalMovement <- "D_Pct"
   TextField "Label_M_V" at 410,388 size 198x16; Text 'M_V'
   Gauge "M_D" at 612,206 size 150x150; CaptionText 'SIMATIC'
      DiagonalMovement <- "D_Pct"
   TextField "Label_M_D" at 612,388 size 198x16; Text 'M_D'
   Gauge "M_Direct" at 814,206 size 150x150; CaptionText 'SIMATIC'
      DirectMovement <- "D_X"
      DirectMovement <- "D_Y"
   TextField "Label_M_Direct" at 814,388 size 198x16; Text 'M_Direct'
   Gauge "E_Range" at 1016,206 size 150x150; CaptionText 'SIMATIC'
      ObjectEnable <- "D_Range"
   TextField "Label_E_Range" at 1016,388 size 198x16; Text 'E_Range'
   Gauge "E_Bit" at 6,408 size 150x150; CaptionText 'SIMATIC'
      ObjectEnable <- "D_En"
   TextField "Label_E_Bit" at 6,590 size 198x16; Text 'E_Bit'
   Gauge "PV_Pct" at 208,408 size 150x150; CaptionText 'SIMATIC'
      ProcessValue <- "D_Pct"
   TextField "Label_PV_Pct" at 208,590 size 198x16; Text 'PV_Pct'
   Gauge "PV_Real" at 410,408 size 150x150; CaptionText 'SIMATIC'
      ProcessValue <- "D_Real"
   TextField "Label_PV_Real" at 410,590 size 198x16; Text 'PV_Real'
   Gauge "PV_Pct_MaxMin" at 612,408 size 150x150; CaptionText 'SIMATIC'
      ProcessValue <- "D_Pct"
      MaximumValue <- "D_Max"
      MinimumValue <- "D_Min"
   TextField "Label_PV_Pct_MaxMin" at 612,590 size 198x16; Text 'PV_Pct_MaxMin'
   IOField "State" at 4,774 size 60x22; FormatPattern 9
      ProcessValue <- "D_State"
   Button "S1" at 70,774 size 40x22; TextOff 'S1'
      on Click: "SetS1"()
   Button "S2" at 114,774 size 40x22; TextOff 'S2'
      on Click: "SetS2"()
   Button "S3" at 158,774 size 40x22; TextOff 'S3'
      on Click: "SetS3"()
   Button "S4" at 202,774 size 40x22; TextOff 'S4'
      on Click: "SetS4"()
   Button "Next" at 1236,774 size 40x22; TextOff 'Next'
      on Click: ActivateScreen("D_Clock_1", 0)

screen "D_GraphicIOField_1" 1280x800
   GraphicIOField "Static" at 6,4 size 60x60
   TextField "Label_Static" at 6,96 size 108x16; Text 'Static'
   GraphicIOField "A_Range" at 118,4 size 60x60
      Appearance <- "D_Range"
   TextField "Label_A_Range" at 118,96 size 108x16; Text 'A_Range'
   GraphicIOField "A_Flash" at 230,4 size 60x60
      Appearance <- "D_Range"
   TextField "Label_A_Flash" at 230,96 size 108x16; Text 'A_Flash'
   GraphicIOField "A_Bit" at 342,4 size 60x60
      Appearance <- "D_Bool"
   TextField "Label_A_Bit" at 342,96 size 108x16; Text 'A_Bit'
   GraphicIOField "A_Bits" at 454,4 size 60x60
      Appearance <- "D_Bits"
   TextField "Label_A_Bits" at 454,96 size 108x16; Text 'A_Bits'
   GraphicIOField "V_Range" at 566,4 size 60x60
      Visibility <- "D_Range"
   TextField "Label_V_Range" at 566,96 size 108x16; Text 'V_Range'
   GraphicIOField "V_Bit" at 678,4 size 60x60
      Visibility <- "D_Vis"
   TextField "Label_V_Bit" at 678,96 size 108x16; Text 'V_Bit'
   GraphicIOField "M_H" at 790,4 size 60x60
      HorizontalMovement <- "D_Pct"
   TextField "Label_M_H" at 790,96 size 108x16; Text 'M_H'
   GraphicIOField "M_V" at 902,4 size 60x60
      VerticalMovement <- "D_Pct"
   TextField "Label_M_V" at 902,96 size 108x16; Text 'M_V'
   GraphicIOField "M_D" at 1014,4 size 60x60
      DiagonalMovement <- "D_Pct"
   TextField "Label_M_D" at 1014,96 size 108x16; Text 'M_D'
   GraphicIOField "M_Direct" at 1126,4 size 60x60
      DirectMovement <- "D_X"
      DirectMovement <- "D_Y"
   TextField "Label_M_Direct" at 1126,96 size 108x16; Text 'M_Direct'
   GraphicIOField "E_Range" at 6,116 size 60x60
      ObjectEnable <- "D_Range"
   TextField "Label_E_Range" at 6,208 size 108x16; Text 'E_Range'
   GraphicIOField "E_Bit" at 118,116 size 60x60
      ObjectEnable <- "D_En"
   TextField "Label_E_Bit" at 118,208 size 108x16; Text 'E_Bit'
   IOField "State" at 4,774 size 60x22; FormatPattern 9
      ProcessValue <- "D_State"
   Button "S1" at 70,774 size 40x22; TextOff 'S1'
      on Click: "SetS1"()
   Button "S2" at 114,774 size 40x22; TextOff 'S2'
      on Click: "SetS2"()
   Button "S3" at 158,774 size 40x22; TextOff 'S3'
      on Click: "SetS3"()
   Button "S4" at 202,774 size 40x22; TextOff 'S4'
      on Click: "SetS4"()
   Button "Next" at 1236,774 size 40x22; TextOff 'Next'
      on Click: ActivateScreen("D_DateTimeField_1", 0)

screen "D_GraphicView_1" 1280x800
   GraphicView "Static" at 6,4 size 100x60
   TextField "Label_Static" at 6,96 size 148x16; Text 'Static'
   GraphicView "A_Range" at 158,4 size 100x60
      Appearance <- "D_Range"
   TextField "Label_A_Range" at 158,96 size 148x16; Text 'A_Range'
   GraphicView "A_Flash" at 310,4 size 100x60
      Appearance <- "D_Range"
   TextField "Label_A_Flash" at 310,96 size 148x16; Text 'A_Flash'
   GraphicView "A_Bit" at 462,4 size 100x60
      Appearance <- "D_Bool"
   TextField "Label_A_Bit" at 462,96 size 148x16; Text 'A_Bit'
   GraphicView "A_Bits" at 614,4 size 100x60
      Appearance <- "D_Bits"
   TextField "Label_A_Bits" at 614,96 size 148x16; Text 'A_Bits'
   GraphicView "V_Range" at 766,4 size 100x60
      Visibility <- "D_Range"
   TextField "Label_V_Range" at 766,96 size 148x16; Text 'V_Range'
   GraphicView "V_Bit" at 918,4 size 100x60
      Visibility <- "D_Vis"
   TextField "Label_V_Bit" at 918,96 size 148x16; Text 'V_Bit'
   GraphicView "M_H" at 1070,4 size 100x60
      HorizontalMovement <- "D_Pct"
   TextField "Label_M_H" at 1070,96 size 148x16; Text 'M_H'
   GraphicView "M_V" at 6,116 size 100x60
      VerticalMovement <- "D_Pct"
   TextField "Label_M_V" at 6,208 size 148x16; Text 'M_V'
   GraphicView "M_D" at 158,116 size 100x60
      DiagonalMovement <- "D_Pct"
   TextField "Label_M_D" at 158,208 size 148x16; Text 'M_D'
   GraphicView "M_Direct" at 310,116 size 100x60
      DirectMovement <- "D_X"
      DirectMovement <- "D_Y"
   TextField "Label_M_Direct" at 310,208 size 148x16; Text 'M_Direct'
   GraphicView "E_Range" at 462,116 size 100x60
      ObjectEnable <- "D_Range"
   TextField "Label_E_Range" at 462,208 size 148x16; Text 'E_Range'
   GraphicView "E_Bit" at 614,116 size 100x60
      ObjectEnable <- "D_En"
   TextField "Label_E_Bit" at 614,208 size 148x16; Text 'E_Bit'
   IOField "State" at 4,774 size 60x22; FormatPattern 9
      ProcessValue <- "D_State"
   Button "S1" at 70,774 size 40x22; TextOff 'S1'
      on Click: "SetS1"()
   Button "S2" at 114,774 size 40x22; TextOff 'S2'
      on Click: "SetS2"()
   Button "S3" at 158,774 size 40x22; TextOff 'S3'
      on Click: "SetS3"()
   Button "S4" at 202,774 size 40x22; TextOff 'S4'
      on Click: "SetS4"()
   Button "Next" at 1236,774 size 40x22; TextOff 'Next'
      on Click: ActivateScreen("D_IOField_1", 0)

screen "D_IOField_1" 1280x800
   IOField "Static" at 6,4 size 100x30
   TextField "Label_Static" at 6,66 size 148x16; Text 'Static'
   IOField "A_Range" at 158,4 size 100x30
      Appearance <- "D_Range"
   TextField "Label_A_Range" at 158,66 size 148x16; Text 'A_Range'
   IOField "A_Flash" at 310,4 size 100x30
      Appearance <- "D_Range"
   TextField "Label_A_Flash" at 310,66 size 148x16; Text 'A_Flash'
   IOField "A_Bit" at 462,4 size 100x30
      Appearance <- "D_Bool"
   TextField "Label_A_Bit" at 462,66 size 148x16; Text 'A_Bit'
   IOField "A_Bits" at 614,4 size 100x30
      Appearance <- "D_Bits"
   TextField "Label_A_Bits" at 614,66 size 148x16; Text 'A_Bits'
   IOField "V_Range" at 766,4 size 100x30
      Visibility <- "D_Range"
   TextField "Label_V_Range" at 766,66 size 148x16; Text 'V_Range'
   IOField "V_Bit" at 918,4 size 100x30
      Visibility <- "D_Vis"
   TextField "Label_V_Bit" at 918,66 size 148x16; Text 'V_Bit'
   IOField "M_H" at 1070,4 size 100x30
      HorizontalMovement <- "D_Pct"
   TextField "Label_M_H" at 1070,66 size 148x16; Text 'M_H'
   IOField "M_V" at 6,86 size 100x30
      VerticalMovement <- "D_Pct"
   TextField "Label_M_V" at 6,148 size 148x16; Text 'M_V'
   IOField "M_D" at 158,86 size 100x30
      DiagonalMovement <- "D_Pct"
   TextField "Label_M_D" at 158,148 size 148x16; Text 'M_D'
   IOField "M_Direct" at 310,86 size 100x30
      DirectMovement <- "D_X"
      DirectMovement <- "D_Y"
   TextField "Label_M_Direct" at 310,148 size 148x16; Text 'M_Direct'
   IOField "E_Range" at 462,86 size 100x30
      ObjectEnable <- "D_Range"
   TextField "Label_E_Range" at 462,148 size 148x16; Text 'E_Range'
   IOField "E_Bit" at 614,86 size 100x30
      ObjectEnable <- "D_En"
   TextField "Label_E_Bit" at 614,148 size 148x16; Text 'E_Bit'
   IOField "PV_SInt" at 766,86 size 100x30; FormatPattern s999
      ProcessValue <- "D_SInt"
   TextField "Label_PV_SInt" at 766,148 size 148x16; Text 'PV_SInt'
   IOField "PV_Int" at 918,86 size 100x30; FormatPattern s99999
      ProcessValue <- "D_Int"
   TextField "Label_PV_Int" at 918,148 size 148x16; Text 'PV_Int'
   IOField "PV_DInt" at 1070,86 size 100x30; FormatPattern s9999999999
      ProcessValue <- "D_DInt"
   TextField "Label_PV_DInt" at 1070,148 size 148x16; Text 'PV_DInt'
   IOField "PV_USInt" at 6,168 size 100x30; FormatPattern 999
      ProcessValue <- "D_USInt"
   TextField "Label_PV_USInt" at 6,230 size 148x16; Text 'PV_USInt'
   IOField "PV_UInt" at 158,168 size 100x30; FormatPattern 99999
      ProcessValue <- "D_UInt"
   TextField "Label_PV_UInt" at 158,230 size 148x16; Text 'PV_UInt'
   IOField "PV_UDInt" at 310,168 size 100x30; FormatPattern 9999999999
      ProcessValue <- "D_UDInt"
   TextField "Label_PV_UDInt" at 310,230 size 148x16; Text 'PV_UDInt'
   IOField "PV_Real" at 462,168 size 100x30
      ProcessValue <- "D_Real"
   TextField "Label_PV_Real" at 462,230 size 148x16; Text 'PV_Real'
   IOField "PV_LReal" at 614,168 size 100x30
      ProcessValue <- "D_LReal"
   TextField "Label_PV_LReal" at 614,230 size 148x16; Text 'PV_LReal'
   IOField "PV_String" at 766,168 size 100x30
      ProcessValue <- "D_String"
   TextField "Label_PV_String" at 766,230 size 148x16; Text 'PV_String'
   IOField "PV_Int_Shift2" at 918,168 size 100x30; FormatPattern s99999
      ProcessValue <- "D_Int"
   TextField "Label_PV_Int_Shift2" at 918,230 size 148x16; Text 'PV_Int_Shift2'
   IOField "PV_Int_s999999" at 1070,168 size 100x30; FormatPattern s999999
      ProcessValue <- "D_Int"
   TextField "Label_PV_Int_s999999" at 1070,230 size 148x16; Text 'PV_Int_s999999'
   IOField "PV_Real_s9999_99" at 6,250 size 100x30; FormatPattern s9999.99
      ProcessValue <- "D_Real"
   TextField "Label_PV_Real_s9999_99" at 6,312 size 148x16; Text 'PV_Real_s9999_99'
   IOField "PV_Int_Output" at 158,250 size 100x30; FormatPattern s99999
      ProcessValue <- "D_Int"
   TextField "Label_PV_Int_Output" at 158,312 size 148x16; Text 'PV_Int_Output'
   IOField "PV_Int_s99" at 310,250 size 100x30; FormatPattern s99
      ProcessValue <- "D_Int"
   TextField "Label_PV_Int_s99" at 310,312 size 148x16; Text 'PV_Int_s99'
   IOField "State" at 4,774 size 60x22; FormatPattern 9
      ProcessValue <- "D_State"
   Button "S1" at 70,774 size 40x22; TextOff 'S1'
      on Click: "SetS1"()
   Button "S2" at 114,774 size 40x22; TextOff 'S2'
      on Click: "SetS2"()
   Button "S3" at 158,774 size 40x22; TextOff 'S3'
      on Click: "SetS3"()
   Button "S4" at 202,774 size 40x22; TextOff 'S4'
      on Click: "SetS4"()
   Button "Next" at 1236,774 size 40x22; TextOff 'Next'
      on Click: ActivateScreen("D_Button_1", 0)

screen "D_Line_1" 1280x800
   TextField "Label_Static" at 6,86 size 148x16; Text 'Static'
   Line "A_Range" at 158,4 size 100x50
      Appearance <- "D_Range"
   TextField "Label_A_Range" at 158,86 size 148x16; Text 'A_Range'
   Line "A_Flash" at 310,4 size 100x50
      Appearance <- "D_Range"
   TextField "Label_A_Flash" at 310,86 size 148x16; Text 'A_Flash'
   Line "A_Bit" at 462,4 size 100x50
      Appearance <- "D_Bool"
   TextField "Label_A_Bit" at 462,86 size 148x16; Text 'A_Bit'
   Line "A_Bits" at 614,4 size 100x50
      Appearance <- "D_Bits"
   TextField "Label_A_Bits" at 614,86 size 148x16; Text 'A_Bits'
   Line "V_Range" at 766,4 size 100x50
      Visibility <- "D_Range"
   TextField "Label_V_Range" at 766,86 size 148x16; Text 'V_Range'
   Line "V_Bit" at 918,4 size 100x50
      Visibility <- "D_Vis"
   TextField "Label_V_Bit" at 918,86 size 148x16; Text 'V_Bit'
   Line "M_H" at 1070,4 size 100x50
      HorizontalMovement <- "D_Pct"
   TextField "Label_M_H" at 1070,86 size 148x16; Text 'M_H'
   Line "M_V" at 6,106 size 100x50
      VerticalMovement <- "D_Pct"
   TextField "Label_M_V" at 6,188 size 148x16; Text 'M_V'
   Line "M_D" at 158,106 size 100x50
      DiagonalMovement <- "D_Pct"
   TextField "Label_M_D" at 158,188 size 148x16; Text 'M_D'
   Line "M_Direct" at 310,106 size 100x50
      DirectMovement <- "D_X"
      DirectMovement <- "D_Y"
   TextField "Label_M_Direct" at 310,188 size 148x16; Text 'M_Direct'
   Line "E_Range" at 462,106 size 100x50
      ObjectEnable <- "D_Range"
   TextField "Label_E_Range" at 462,188 size 148x16; Text 'E_Range'
   Line "E_Bit" at 614,106 size 100x50
      ObjectEnable <- "D_En"
   TextField "Label_E_Bit" at 614,188 size 148x16; Text 'E_Bit'
   IOField "State" at 4,774 size 60x22; FormatPattern 9
      ProcessValue <- "D_State"
   Button "S1" at 70,774 size 40x22; TextOff 'S1'
      on Click: "SetS1"()
   Button "S2" at 114,774 size 40x22; TextOff 'S2'
      on Click: "SetS2"()
   Button "S3" at 158,774 size 40x22; TextOff 'S3'
      on Click: "SetS3"()
   Button "S4" at 202,774 size 40x22; TextOff 'S4'
      on Click: "SetS4"()
   Button "Next" at 1236,774 size 40x22; TextOff 'Next'
      on Click: ActivateScreen("D_Polyline_1", 0)

screen "D_Polygon_1" 1280x800
   TextField "Label_Static" at 6,86 size 148x16; Text 'Static'
   Polygon "A_Range" at 158,4 size 100x50
      Appearance <- "D_Range"
   TextField "Label_A_Range" at 158,86 size 148x16; Text 'A_Range'
   Polygon "A_Flash" at 310,4 size 100x50
      Appearance <- "D_Range"
   TextField "Label_A_Flash" at 310,86 size 148x16; Text 'A_Flash'
   Polygon "A_Bit" at 462,4 size 100x50
      Appearance <- "D_Bool"
   TextField "Label_A_Bit" at 462,86 size 148x16; Text 'A_Bit'
   Polygon "A_Bits" at 614,4 size 100x50
      Appearance <- "D_Bits"
   TextField "Label_A_Bits" at 614,86 size 148x16; Text 'A_Bits'
   Polygon "V_Range" at 766,4 size 100x50
      Visibility <- "D_Range"
   TextField "Label_V_Range" at 766,86 size 148x16; Text 'V_Range'
   Polygon "V_Bit" at 918,4 size 100x50
      Visibility <- "D_Vis"
   TextField "Label_V_Bit" at 918,86 size 148x16; Text 'V_Bit'
   Polygon "M_H" at 1070,4 size 100x50
      HorizontalMovement <- "D_Pct"
   TextField "Label_M_H" at 1070,86 size 148x16; Text 'M_H'
   Polygon "M_V" at 6,106 size 100x50
      VerticalMovement <- "D_Pct"
   TextField "Label_M_V" at 6,188 size 148x16; Text 'M_V'
   Polygon "M_D" at 158,106 size 100x50
      DiagonalMovement <- "D_Pct"
   TextField "Label_M_D" at 158,188 size 148x16; Text 'M_D'
   Polygon "M_Direct" at 310,106 size 100x50
      DirectMovement <- "D_X"
      DirectMovement <- "D_Y"
   TextField "Label_M_Direct" at 310,188 size 148x16; Text 'M_Direct'
   Polygon "E_Range" at 462,106 size 100x50
      ObjectEnable <- "D_Range"
   TextField "Label_E_Range" at 462,188 size 148x16; Text 'E_Range'
   Polygon "E_Bit" at 614,106 size 100x50
      ObjectEnable <- "D_En"
   TextField "Label_E_Bit" at 614,188 size 148x16; Text 'E_Bit'
   IOField "State" at 4,774 size 60x22; FormatPattern 9
      ProcessValue <- "D_State"
   Button "S1" at 70,774 size 40x22; TextOff 'S1'
      on Click: "SetS1"()
   Button "S2" at 114,774 size 40x22; TextOff 'S2'
      on Click: "SetS2"()
   Button "S3" at 158,774 size 40x22; TextOff 'S3'
      on Click: "SetS3"()
   Button "S4" at 202,774 size 40x22; TextOff 'S4'
      on Click: "SetS4"()
   Button "Next" at 1236,774 size 40x22; TextOff 'Next'
      on Click: ActivateScreen("D_Ellipse_1", 0)

screen "D_Polyline_1" 1280x800
   TextField "Label_Static" at 6,86 size 148x16; Text 'Static'
   Polyline "A_Range" at 158,4 size 100x50
      Appearance <- "D_Range"
   TextField "Label_A_Range" at 158,86 size 148x16; Text 'A_Range'
   Polyline "A_Flash" at 310,4 size 100x50
      Appearance <- "D_Range"
   TextField "Label_A_Flash" at 310,86 size 148x16; Text 'A_Flash'
   Polyline "A_Bit" at 462,4 size 100x50
      Appearance <- "D_Bool"
   TextField "Label_A_Bit" at 462,86 size 148x16; Text 'A_Bit'
   Polyline "A_Bits" at 614,4 size 100x50
      Appearance <- "D_Bits"
   TextField "Label_A_Bits" at 614,86 size 148x16; Text 'A_Bits'
   Polyline "V_Range" at 766,4 size 100x50
      Visibility <- "D_Range"
   TextField "Label_V_Range" at 766,86 size 148x16; Text 'V_Range'
   Polyline "V_Bit" at 918,4 size 100x50
      Visibility <- "D_Vis"
   TextField "Label_V_Bit" at 918,86 size 148x16; Text 'V_Bit'
   Polyline "M_H" at 1070,4 size 100x50
      HorizontalMovement <- "D_Pct"
   TextField "Label_M_H" at 1070,86 size 148x16; Text 'M_H'
   Polyline "M_V" at 6,106 size 100x50
      VerticalMovement <- "D_Pct"
   TextField "Label_M_V" at 6,188 size 148x16; Text 'M_V'
   Polyline "M_D" at 158,106 size 100x50
      DiagonalMovement <- "D_Pct"
   TextField "Label_M_D" at 158,188 size 148x16; Text 'M_D'
   Polyline "M_Direct" at 310,106 size 100x50
      DirectMovement <- "D_X"
      DirectMovement <- "D_Y"
   TextField "Label_M_Direct" at 310,188 size 148x16; Text 'M_Direct'
   Polyline "E_Range" at 462,106 size 100x50
      ObjectEnable <- "D_Range"
   TextField "Label_E_Range" at 462,188 size 148x16; Text 'E_Range'
   Polyline "E_Bit" at 614,106 size 100x50
      ObjectEnable <- "D_En"
   TextField "Label_E_Bit" at 614,188 size 148x16; Text 'E_Bit'
   IOField "State" at 4,774 size 60x22; FormatPattern 9
      ProcessValue <- "D_State"
   Button "S1" at 70,774 size 40x22; TextOff 'S1'
      on Click: "SetS1"()
   Button "S2" at 114,774 size 40x22; TextOff 'S2'
      on Click: "SetS2"()
   Button "S3" at 158,774 size 40x22; TextOff 'S3'
      on Click: "SetS3"()
   Button "S4" at 202,774 size 40x22; TextOff 'S4'
      on Click: "SetS4"()
   Button "Next" at 1236,774 size 40x22; TextOff 'Next'
      on Click: ActivateScreen("D_Polygon_1", 0)

